REGION Network 5: Tempo total do sinal da fabrica
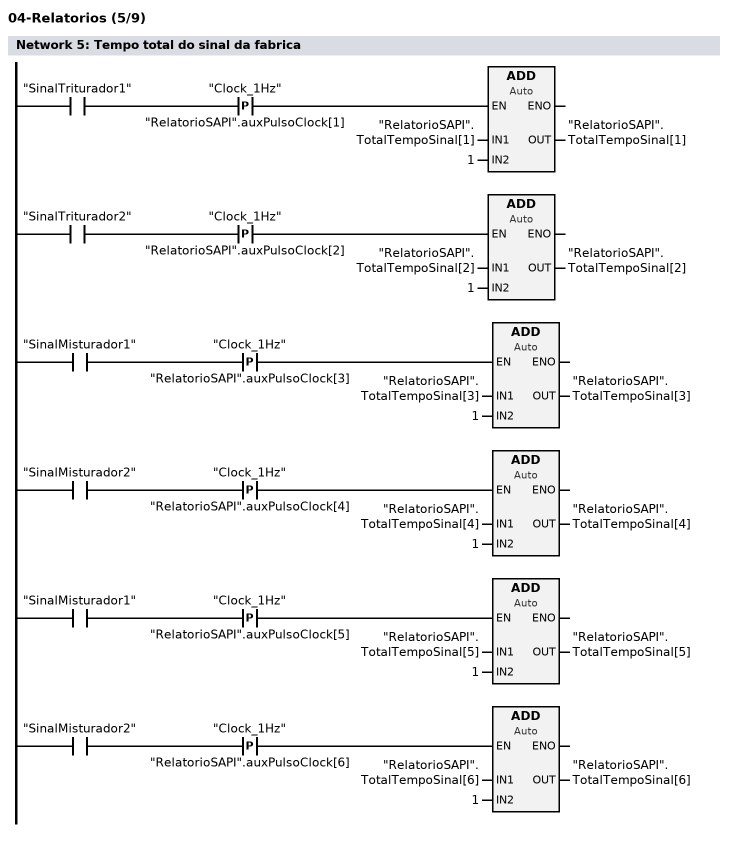
   RUNG wire#powerrail
      Contact( "SinalTriturador1" )
      P_Contact(operand := "Clock_1Hz", bit := "RelatorioSAPI".auxPulsoClock[1])
      Add(in1 := "RelatorioSAPI".TotalTempoSinal[1], in2 := 1, out => "RelatorioSAPI".TotalTempoSinal[1])
   END_RUNG
   RUNG wire#powerrail
      Contact( "SinalTriturador2" )
      P_Contact(operand := "Clock_1Hz", bit := "RelatorioSAPI".auxPulsoClock[2])
      Add(in1 := "RelatorioSAPI".TotalTempoSinal[2], in2 := 1, out => "RelatorioSAPI".TotalTempoSinal[2])
   END_RUNG
   RUNG wire#powerrail
      Contact( "SinalMisturador1" )
      P_Contact(operand := "Clock_1Hz", bit := "RelatorioSAPI".auxPulsoClock[3])
      Add(in1 := "RelatorioSAPI".TotalTempoSinal[3], in2 := 1, out => "RelatorioSAPI".TotalTempoSinal[3])
   END_RUNG
   RUNG wire#powerrail
      Contact( "SinalMisturador2" )
      P_Contact(operand := "Clock_1Hz", bit := "RelatorioSAPI".auxPulsoClock[4])
      Add(in1 := "RelatorioSAPI".TotalTempoSinal[4], in2 := 1, out => "RelatorioSAPI".TotalTempoSinal[4])
   END_RUNG
   RUNG wire#powerrail
      Contact( "SinalMisturador1" )
      P_Contact(operand := "Clock_1Hz", bit := "RelatorioSAPI".auxPulsoClock[5])
      Add(in1 := "RelatorioSAPI".TotalTempoSinal[5], in2 := 1, out => "RelatorioSAPI".TotalTempoSinal[5])
   END_RUNG
   RUNG wire#powerrail
      Contact( "SinalMisturador2" )
      P_Contact(operand := "Clock_1Hz", bit := "RelatorioSAPI".auxPulsoClock[6])
      Add(in1 := "RelatorioSAPI".TotalTempoSinal[6], in2 := 1, out => "RelatorioSAPI".TotalTempoSinal[6])
   END_RUNG
   // the same network as SCL:
   #_w1 := "SinalTriturador1" AND "Clock_1Hz" AND NOT "RelatorioSAPI".auxPulsoClock[1];   // rising edge of "Clock_1Hz"
   "RelatorioSAPI".auxPulsoClock[1] := "Clock_1Hz";
   IF #_w1 THEN "RelatorioSAPI".TotalTempoSinal[1] := "RelatorioSAPI".TotalTempoSinal[1] + 1; END_IF;
   #_w2 := "SinalTriturador2" AND "Clock_1Hz" AND NOT "RelatorioSAPI".auxPulsoClock[2];   // rising edge of "Clock_1Hz"
   "RelatorioSAPI".auxPulsoClock[2] := "Clock_1Hz";
   IF #_w2 THEN "RelatorioSAPI".TotalTempoSinal[2] := "RelatorioSAPI".TotalTempoSinal[2] + 1; END_IF;
   #_w3 := "SinalMisturador1" AND "Clock_1Hz" AND NOT "RelatorioSAPI".auxPulsoClock[3];   // rising edge of "Clock_1Hz"
   "RelatorioSAPI".auxPulsoClock[3] := "Clock_1Hz";
   IF #_w3 THEN "RelatorioSAPI".TotalTempoSinal[3] := "RelatorioSAPI".TotalTempoSinal[3] + 1; END_IF;
   #_w4 := "SinalMisturador2" AND "Clock_1Hz" AND NOT "RelatorioSAPI".auxPulsoClock[4];   // rising edge of "Clock_1Hz"
   "RelatorioSAPI".auxPulsoClock[4] := "Clock_1Hz";
   IF #_w4 THEN "RelatorioSAPI".TotalTempoSinal[4] := "RelatorioSAPI".TotalTempoSinal[4] + 1; END_IF;
   #_w5 := "SinalMisturador1" AND "Clock_1Hz" AND NOT "RelatorioSAPI".auxPulsoClock[5];   // rising edge of "Clock_1Hz"
   "RelatorioSAPI".auxPulsoClock[5] := "Clock_1Hz";
   IF #_w5 THEN "RelatorioSAPI".TotalTempoSinal[5] := "RelatorioSAPI".TotalTempoSinal[5] + 1; END_IF;
   #_w6 := "SinalMisturador2" AND "Clock_1Hz" AND NOT "RelatorioSAPI".auxPulsoClock[6];   // rising edge of "Clock_1Hz"
   "RelatorioSAPI".auxPulsoClock[6] := "Clock_1Hz";
   IF #_w6 THEN "RelatorioSAPI".TotalTempoSinal[6] := "RelatorioSAPI".TotalTempoSinal[6] + 1; END_IF;
END_REGION

REGION Network 6: Quantidade acionamentos sinal fabrica
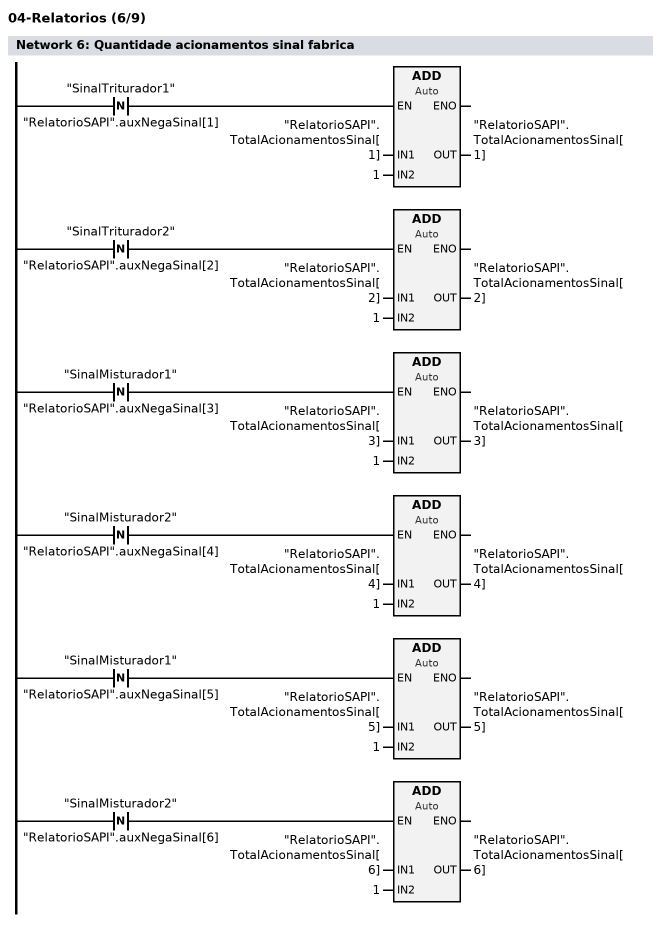
   RUNG wire#powerrail
      N_Contact(operand := "SinalTriturador1", bit := "RelatorioSAPI".auxNegaSinal[1])
      Add(in1 := "RelatorioSAPI".TotalAcionamentosSinal[1], in2 := 1, out => "RelatorioSAPI".TotalAcionamentosSinal[1])
   END_RUNG
   RUNG wire#powerrail
      N_Contact(operand := "SinalTriturador2", bit := "RelatorioSAPI".auxNegaSinal[2])
      Add(in1 := "RelatorioSAPI".TotalAcionamentosSinal[2], in2 := 1, out => "RelatorioSAPI".TotalAcionamentosSinal[2])
   END_RUNG
   RUNG wire#powerrail
      N_Contact(operand := "SinalMisturador1", bit := "RelatorioSAPI".auxNegaSinal[3])
      Add(in1 := "RelatorioSAPI".TotalAcionamentosSinal[3], in2 := 1, out => "RelatorioSAPI".TotalAcionamentosSinal[3])
   END_RUNG
   RUNG wire#powerrail
      N_Contact(operand := "SinalMisturador2", bit := "RelatorioSAPI".auxNegaSinal[4])
      Add(in1 := "RelatorioSAPI".TotalAcionamentosSinal[4], in2 := 1, out => "RelatorioSAPI".TotalAcionamentosSinal[4])
   END_RUNG
   RUNG wire#powerrail
      N_Contact(operand := "SinalMisturador1", bit := "RelatorioSAPI".auxNegaSinal[5])
      Add(in1 := "RelatorioSAPI".TotalAcionamentosSinal[5], in2 := 1, out => "RelatorioSAPI".TotalAcionamentosSinal[5])
   END_RUNG
   RUNG wire#powerrail
      N_Contact(operand := "SinalMisturador2", bit := "RelatorioSAPI".auxNegaSinal[6])
      Add(in1 := "RelatorioSAPI".TotalAcionamentosSinal[6], in2 := 1, out => "RelatorioSAPI".TotalAcionamentosSinal[6])
   END_RUNG
   // the same network as SCL:
   #_w1 := NOT "SinalTriturador1" AND "RelatorioSAPI".auxNegaSinal[1];   // falling edge of "SinalTriturador1"
   "RelatorioSAPI".auxNegaSinal[1] := "SinalTriturador1";
   IF #_w1 THEN
       "RelatorioSAPI".TotalAcionamentosSinal[1] := "RelatorioSAPI".TotalAcionamentosSinal[1] + 1;
   END_IF;
   #_w2 := NOT "SinalTriturador2" AND "RelatorioSAPI".auxNegaSinal[2];   // falling edge of "SinalTriturador2"
   "RelatorioSAPI".auxNegaSinal[2] := "SinalTriturador2";
   IF #_w2 THEN
       "RelatorioSAPI".TotalAcionamentosSinal[2] := "RelatorioSAPI".TotalAcionamentosSinal[2] + 1;
   END_IF;
   #_w3 := NOT "SinalMisturador1" AND "RelatorioSAPI".auxNegaSinal[3];   // falling edge of "SinalMisturador1"
   "RelatorioSAPI".auxNegaSinal[3] := "SinalMisturador1";
   IF #_w3 THEN
       "RelatorioSAPI".TotalAcionamentosSinal[3] := "RelatorioSAPI".TotalAcionamentosSinal[3] + 1;
   END_IF;
   #_w4 := NOT "SinalMisturador2" AND "RelatorioSAPI".auxNegaSinal[4];   // falling edge of "SinalMisturador2"
   "RelatorioSAPI".auxNegaSinal[4] := "SinalMisturador2";
   IF #_w4 THEN
       "RelatorioSAPI".TotalAcionamentosSinal[4] := "RelatorioSAPI".TotalAcionamentosSinal[4] + 1;
   END_IF;
   #_w5 := NOT "SinalMisturador1" AND "RelatorioSAPI".auxNegaSinal[5];   // falling edge of "SinalMisturador1"
   "RelatorioSAPI".auxNegaSinal[5] := "SinalMisturador1";
   IF #_w5 THEN
       "RelatorioSAPI".TotalAcionamentosSinal[5] := "RelatorioSAPI".TotalAcionamentosSinal[5] + 1;
   END_IF;
   #_w6 := NOT "SinalMisturador2" AND "RelatorioSAPI".auxNegaSinal[6];   // falling edge of "SinalMisturador2"
   "RelatorioSAPI".auxNegaSinal[6] := "SinalMisturador2";
   IF #_w6 THEN
       "RelatorioSAPI".TotalAcionamentosSinal[6] := "RelatorioSAPI".TotalAcionamentosSinal[6] + 1;
   END_IF;
END_REGION

REGION Network 7: Quantidade acionamentos bombas
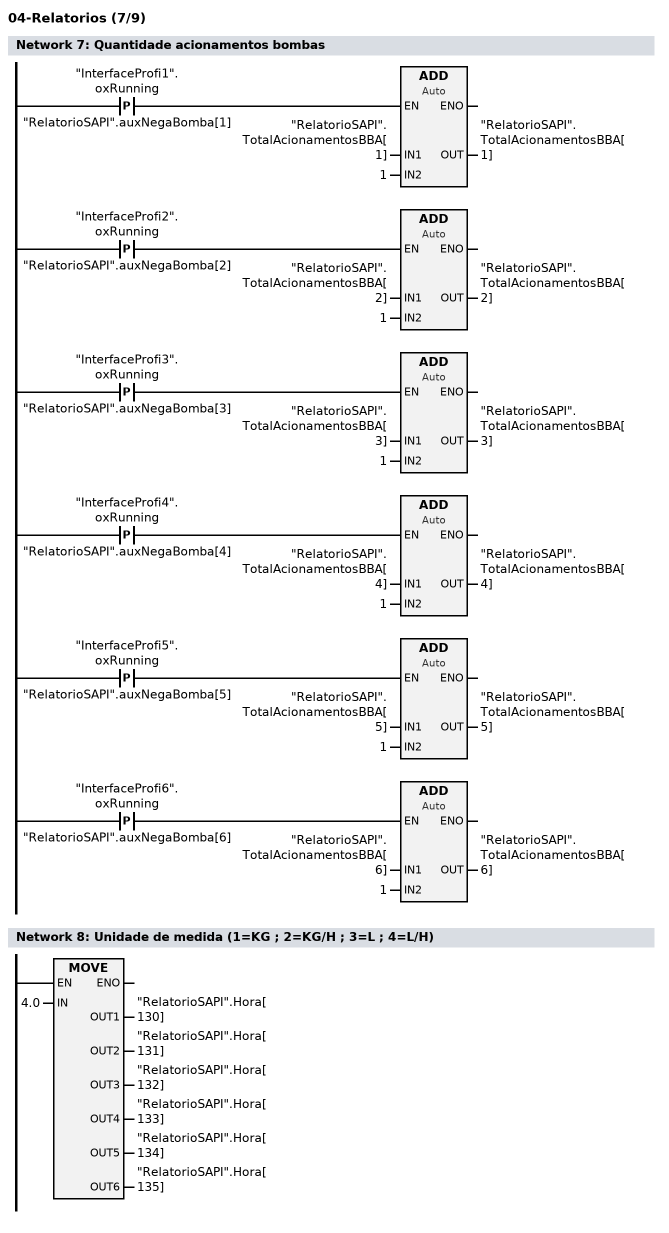
   RUNG wire#powerrail
      P_Contact(operand := "InterfaceProfi1".oxRunning, bit := "RelatorioSAPI".auxNegaBomba[1])
      Add(in1 := "RelatorioSAPI".TotalAcionamentosBBA[1], in2 := 1, out => "RelatorioSAPI".TotalAcionamentosBBA[1])
   END_RUNG
   RUNG wire#powerrail
      P_Contact(operand := "InterfaceProfi2".oxRunning, bit := "RelatorioSAPI".auxNegaBomba[2])
      Add(in1 := "RelatorioSAPI".TotalAcionamentosBBA[2], in2 := 1, out => "RelatorioSAPI".TotalAcionamentosBBA[2])
   END_RUNG
   RUNG wire#powerrail
      P_Contact(operand := "InterfaceProfi3".oxRunning, bit := "RelatorioSAPI".auxNegaBomba[3])
      Add(in1 := "RelatorioSAPI".TotalAcionamentosBBA[3], in2 := 1, out => "RelatorioSAPI".TotalAcionamentosBBA[3])
   END_RUNG
   RUNG wire#powerrail
      P_Contact(operand := "InterfaceProfi4".oxRunning, bit := "RelatorioSAPI".auxNegaBomba[4])
      Add(in1 := "RelatorioSAPI".TotalAcionamentosBBA[4], in2 := 1, out => "RelatorioSAPI".TotalAcionamentosBBA[4])
   END_RUNG
   RUNG wire#powerrail
      P_Contact(operand := "InterfaceProfi5".oxRunning, bit := "RelatorioSAPI".auxNegaBomba[5])
      Add(in1 := "RelatorioSAPI".TotalAcionamentosBBA[5], in2 := 1, out => "RelatorioSAPI".TotalAcionamentosBBA[5])
   END_RUNG
   RUNG wire#powerrail
      P_Contact(operand := "InterfaceProfi6".oxRunning, bit := "RelatorioSAPI".auxNegaBomba[6])
      Add(in1 := "RelatorioSAPI".TotalAcionamentosBBA[6], in2 := 1, out => "RelatorioSAPI".TotalAcionamentosBBA[6])
   END_RUNG
   // the same network as SCL:
   #_w1 := "InterfaceProfi1".oxRunning AND NOT "RelatorioSAPI".auxNegaBomba[1];   // rising edge of "InterfaceProfi1".oxRunning
   "RelatorioSAPI".auxNegaBomba[1] := "InterfaceProfi1".oxRunning;
   IF #_w1 THEN
       "RelatorioSAPI".TotalAcionamentosBBA[1] := "RelatorioSAPI".TotalAcionamentosBBA[1] + 1;
   END_IF;
   #_w2 := "InterfaceProfi2".oxRunning AND NOT "RelatorioSAPI".auxNegaBomba[2];   // rising edge of "InterfaceProfi2".oxRunning
   "RelatorioSAPI".auxNegaBomba[2] := "InterfaceProfi2".oxRunning;
   IF #_w2 THEN
       "RelatorioSAPI".TotalAcionamentosBBA[2] := "RelatorioSAPI".TotalAcionamentosBBA[2] + 1;
   END_IF;
   #_w3 := "InterfaceProfi3".oxRunning AND NOT "RelatorioSAPI".auxNegaBomba[3];   // rising edge of "InterfaceProfi3".oxRunning
   "RelatorioSAPI".auxNegaBomba[3] := "InterfaceProfi3".oxRunning;
   IF #_w3 THEN
       "RelatorioSAPI".TotalAcionamentosBBA[3] := "RelatorioSAPI".TotalAcionamentosBBA[3] + 1;
   END_IF;
   #_w4 := "InterfaceProfi4".oxRunning AND NOT "RelatorioSAPI".auxNegaBomba[4];   // rising edge of "InterfaceProfi4".oxRunning
   "RelatorioSAPI".auxNegaBomba[4] := "InterfaceProfi4".oxRunning;
   IF #_w4 THEN
       "RelatorioSAPI".TotalAcionamentosBBA[4] := "RelatorioSAPI".TotalAcionamentosBBA[4] + 1;
   END_IF;
   #_w5 := "InterfaceProfi5".oxRunning AND NOT "RelatorioSAPI".auxNegaBomba[5];   // rising edge of "InterfaceProfi5".oxRunning
   "RelatorioSAPI".auxNegaBomba[5] := "InterfaceProfi5".oxRunning;
   IF #_w5 THEN
       "RelatorioSAPI".TotalAcionamentosBBA[5] := "RelatorioSAPI".TotalAcionamentosBBA[5] + 1;
   END_IF;
   #_w6 := "InterfaceProfi6".oxRunning AND NOT "RelatorioSAPI".auxNegaBomba[6];   // rising edge of "InterfaceProfi6".oxRunning
   "RelatorioSAPI".auxNegaBomba[6] := "InterfaceProfi6".oxRunning;
   IF #_w6 THEN
       "RelatorioSAPI".TotalAcionamentosBBA[6] := "RelatorioSAPI".TotalAcionamentosBBA[6] + 1;
   END_IF;
END_REGION

REGION Network 8: Unidade de medida (1=KG ; 2=KG/H ; 3=L ; 4=L/H)
   RUNG wire#powerrail
      Move(in := 4.0, out1 => "RelatorioSAPI".Hora[130], out2 => "RelatorioSAPI".Hora[131], out3 => "RelatorioSAPI".Hora[132], out4 => "RelatorioSAPI".Hora[133], out5 => "RelatorioSAPI".Hora[134], out6 => "RelatorioSAPI".Hora[135])
   END_RUNG
   // the same network as SCL:
   "RelatorioSAPI".Hora[130] := 4.0;
   "RelatorioSAPI".Hora[131] := 4.0;
   "RelatorioSAPI".Hora[132] := 4.0;
   "RelatorioSAPI".Hora[133] := 4.0;
   "RelatorioSAPI".Hora[134] := 4.0;
   "RelatorioSAPI".Hora[135] := 4.0;
END_REGION

REGION Network 9: NOME DA BOMBA
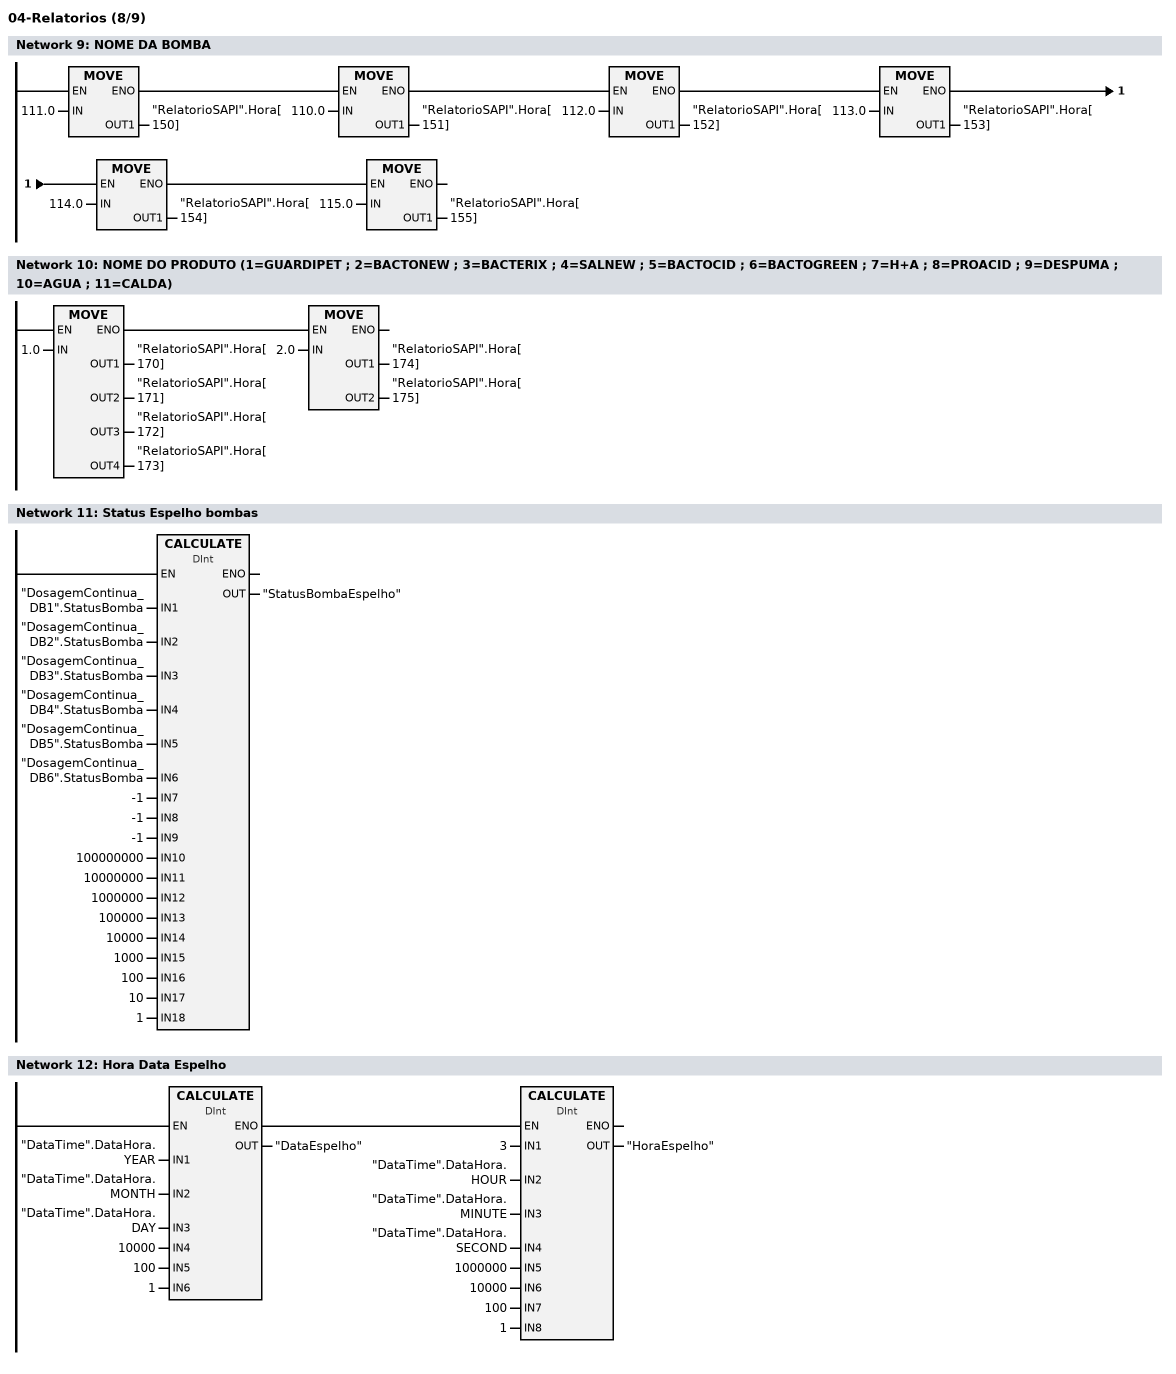
   RUNG wire#powerrail
      Move(in := 111.0, out1 => "RelatorioSAPI".Hora[150])
      Move(in := 110.0, out1 => "RelatorioSAPI".Hora[151])
      Move(in := 112.0, out1 => "RelatorioSAPI".Hora[152])
      Move(in := 113.0, out1 => "RelatorioSAPI".Hora[153])
      Move(in := 114.0, out1 => "RelatorioSAPI".Hora[154])
      Move(in := 115.0, out1 => "RelatorioSAPI".Hora[155])
   END_RUNG
   // the same network as SCL:
   "RelatorioSAPI".Hora[150] := 111.0;
   "RelatorioSAPI".Hora[151] := 110.0;
   "RelatorioSAPI".Hora[152] := 112.0;
   "RelatorioSAPI".Hora[153] := 113.0;
   "RelatorioSAPI".Hora[154] := 114.0;
   "RelatorioSAPI".Hora[155] := 115.0;
END_REGION

REGION Network 10: NOME DO PRODUTO (1=GUARDIPET ; 2=BACTONEW ; 3=BACTERIX ; 4=SALNEW ; 5=BACTOCID ; 6=BACTOGREEN ; 7=H+A ; 8=PROACID ; 9=DESPUMA ; 10=AGUA ; 11=CALDA)
   RUNG wire#powerrail
      Move(in := 1.0, out1 => "RelatorioSAPI".Hora[170], out2 => "RelatorioSAPI".Hora[171], out3 => "RelatorioSAPI".Hora[172], out4 => "RelatorioSAPI".Hora[173])
      Move(in := 2.0, out1 => "RelatorioSAPI".Hora[174], out2 => "RelatorioSAPI".Hora[175])
   END_RUNG
   // the same network as SCL:
   "RelatorioSAPI".Hora[170] := 1.0;
   "RelatorioSAPI".Hora[171] := 1.0;
   "RelatorioSAPI".Hora[172] := 1.0;
   "RelatorioSAPI".Hora[173] := 1.0;
   "RelatorioSAPI".Hora[174] := 2.0;
   "RelatorioSAPI".Hora[175] := 2.0;
END_REGION

REGION Network 11: Status Espelho bombas
   RUNG wire#powerrail
      { S7_Templates := "SrcType := DInt"; S7_Expression := "(((IN18+IN1) * IN10) + ((IN18+IN2) * IN11) + ((IN18+IN3) * IN12) + ((IN18+IN4) * IN13) + ((IN18+IN5) * IN14) + ((IN18+IN6) * IN15) + ((IN18+IN7) * IN16) + ((IN18+IN8) * IN17) + ((IN18+IN9) * IN18))" } Calculate(in1 := "DosagemContinua_DB1".StatusBomba, in2 := "DosagemContinua_DB2".StatusBomba, in3 := "DosagemContinua_DB3".StatusBomba, in4 := "DosagemContinua_DB4".StatusBomba, in5 := "DosagemContinua_DB5".StatusBomba, in6 := "DosagemContinua_DB6".StatusBomba, in7 := -1, in8 := -1, in9 := -1, in10 := 100000000, in11 := 10000000, in12 := 1000000, in13 := 100000, in14 := 10000, in15 := 1000, in16 := 100, in17 := 10, in18 := 1, out => "StatusBombaEspelho")
   END_RUNG
   // the same network as SCL:
   "StatusBombaEspelho" := (((1+"DosagemContinua_DB1".StatusBomba) * 100000000) + ((1+"DosagemContinua_DB2".StatusBomba) * 10000000) + ((1+"DosagemContinua_DB3".StatusBomba) * 1000000) + ((1+"DosagemContinua_DB4".StatusBomba) * 100000) + ((1+"DosagemContinua_DB5".StatusBomba) * 10000) + ((1+"DosagemContinua_DB6".StatusBomba) * 1000) + ((1+(-1)) * 100) + ((1+(-1)) * 10) + ((1+(-1)) * 1));
END_REGION

REGION Network 12: Hora Data Espelho
   RUNG wire#powerrail
      { S7_Templates := "SrcType := DInt"; S7_Expression := "((IN1 * IN4) + (IN2 * IN5) + (IN3 * IN6))" } Calculate(in1 := "DataTime".DataHora.YEAR, in2 := "DataTime".DataHora.MONTH, in3 := "DataTime".DataHora.DAY, in4 := 10000, in5 := 100, in6 := 1, out => "DataEspelho")
      { S7_Templates := "SrcType := DInt"; S7_Expression := "((IN1 * IN5) + (IN2 * IN6) + (IN3 * IN7) + (IN4 * IN8))" } Calculate(in1 := 3, in2 := "DataTime".DataHora.HOUR, in3 := "DataTime".DataHora.MINUTE, in4 := "DataTime".DataHora.SECOND, in5 := 1000000, in6 := 10000, in7 := 100, in8 := 1, out => "HoraEspelho")
   END_RUNG
   // the same network as SCL:
   "DataEspelho" := (("DataTime".DataHora.YEAR * 10000) + ("DataTime".DataHora.MONTH * 100) + ("DataTime".DataHora.DAY * 1));
   "HoraEspelho" := ((3 * 1000000) + ("DataTime".DataHora.HOUR * 10000) + ("DataTime".DataHora.MINUTE * 100) + ("DataTime".DataHora.SECOND * 1));
END_REGION

REGION Network 13: RELATORIO SAPI
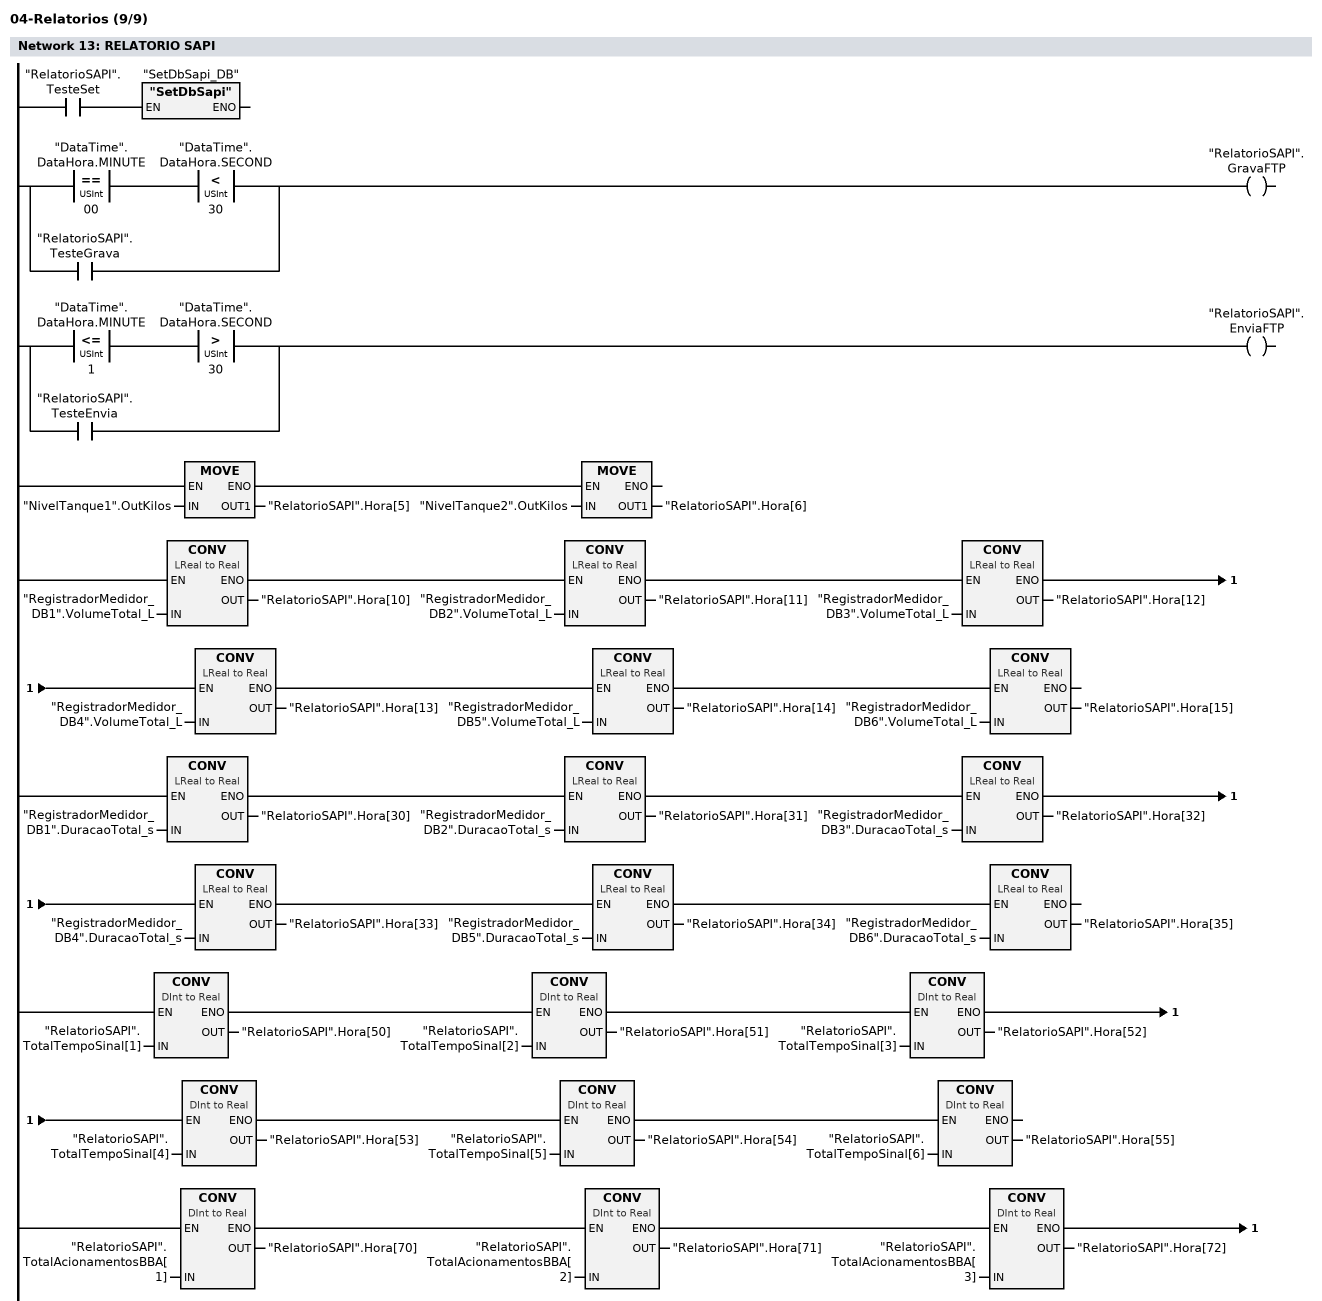
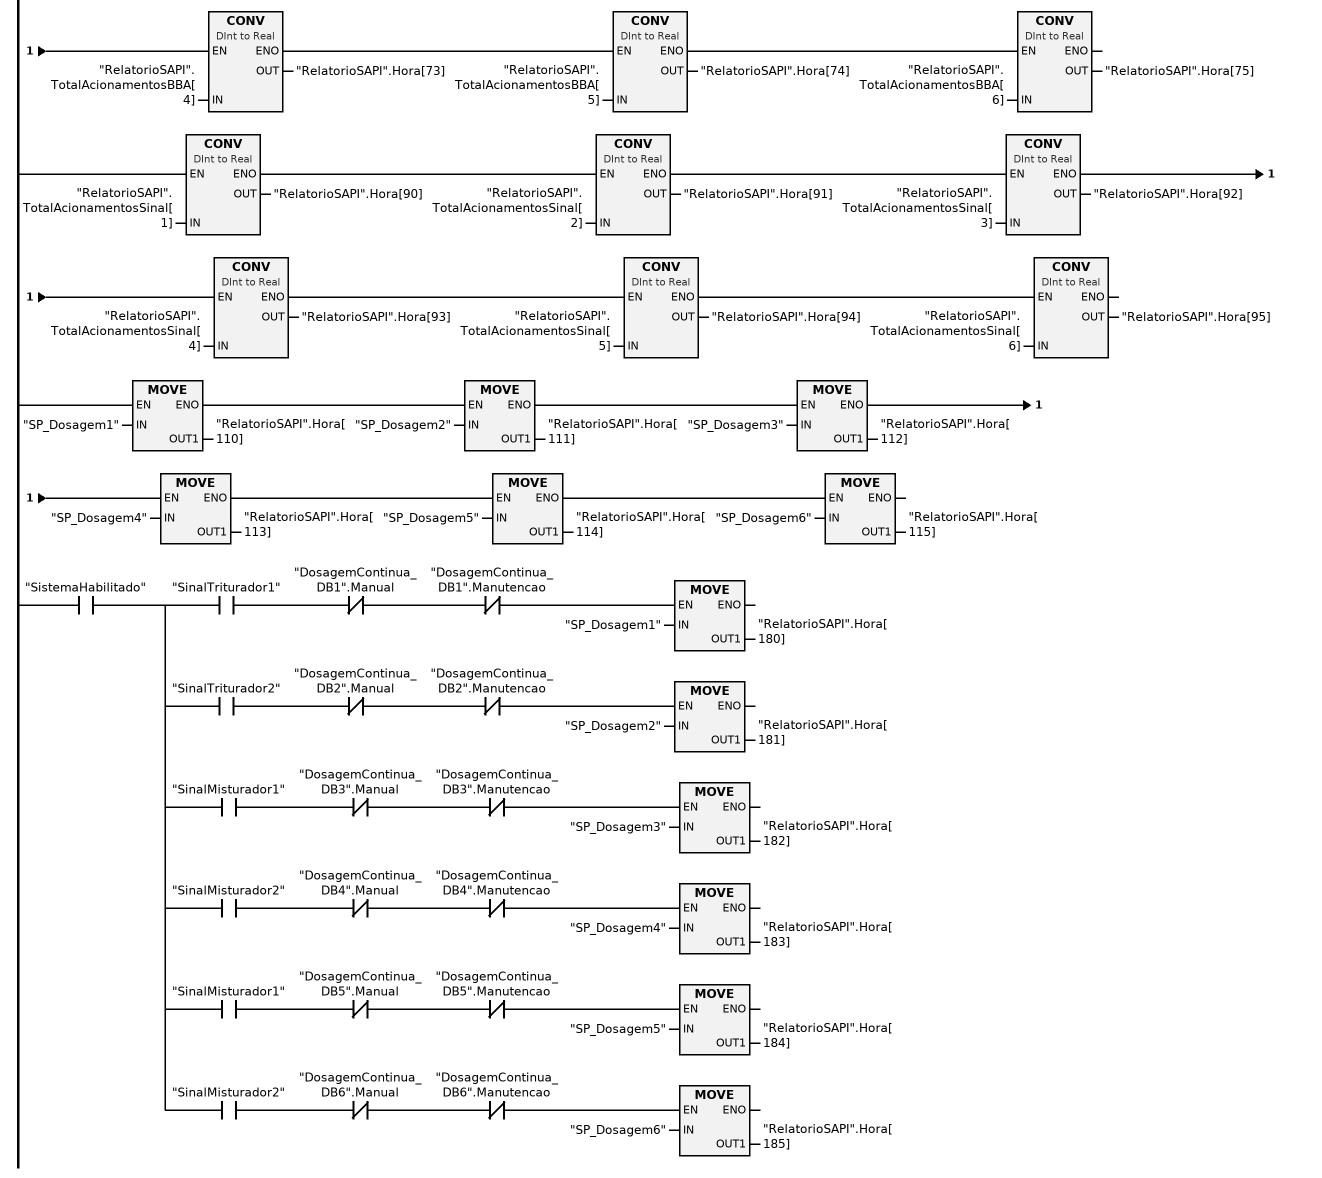
   RUNG wire#powerrail
      Contact( "RelatorioSAPI".TesteSet )
      "SetDbSapi_DB"()
   END_RUNG
   RUNG wire#powerrail
      { S7_Templates := "SrcType := USInt" } EQ_Contact(in1 := "DataTime".DataHora.MINUTE, in2 := 00)
      { S7_Templates := "SrcType := USInt" } LT_Contact(in1 := "DataTime".DataHora.SECOND, in2 := 30)
      wire#w1
      Coil( "RelatorioSAPI".GravaFTP )
   END_RUNG
   RUNG wire#powerrail
      Contact( "RelatorioSAPI".TesteGrava )
   END_RUNG wire#w1
   RUNG wire#powerrail
      { S7_Templates := "SrcType := USInt" } LE_Contact(in1 := "DataTime".DataHora.MINUTE, in2 := 1)
      { S7_Templates := "SrcType := USInt" } GT_Contact(in1 := "DataTime".DataHora.SECOND, in2 := 30)
      wire#w2
      Coil( "RelatorioSAPI".EnviaFTP )
   END_RUNG
   RUNG wire#powerrail
      Contact( "RelatorioSAPI".TesteEnvia )
   END_RUNG wire#w2
   RUNG wire#powerrail
      Move(in := "NivelTanque1".OutKilos, out1 => "RelatorioSAPI".Hora[5])
      Move(in := "NivelTanque2".OutKilos, out1 => "RelatorioSAPI".Hora[6])
   END_RUNG
   RUNG wire#powerrail
      { S7_Templates := "[SrcType := LReal, DestType := Real]" } Convert(in := "RegistradorMedidor_DB1".VolumeTotal_L, out => "RelatorioSAPI".Hora[10])
      { S7_Templates := "[SrcType := LReal, DestType := Real]" } Convert(in := "RegistradorMedidor_DB2".VolumeTotal_L, out => "RelatorioSAPI".Hora[11])
      { S7_Templates := "[SrcType := LReal, DestType := Real]" } Convert(in := "RegistradorMedidor_DB3".VolumeTotal_L, out => "RelatorioSAPI".Hora[12])
      { S7_Templates := "[SrcType := LReal, DestType := Real]" } Convert(in := "RegistradorMedidor_DB4".VolumeTotal_L, out => "RelatorioSAPI".Hora[13])
      { S7_Templates := "[SrcType := LReal, DestType := Real]" } Convert(in := "RegistradorMedidor_DB5".VolumeTotal_L, out => "RelatorioSAPI".Hora[14])
      { S7_Templates := "[SrcType := LReal, DestType := Real]" } Convert(in := "RegistradorMedidor_DB6".VolumeTotal_L, out => "RelatorioSAPI".Hora[15])
   END_RUNG
   RUNG wire#powerrail
      { S7_Templates := "[SrcType := LReal, DestType := Real]" } Convert(in := "RegistradorMedidor_DB1".DuracaoTotal_s, out => "RelatorioSAPI".Hora[30])
      { S7_Templates := "[SrcType := LReal, DestType := Real]" } Convert(in := "RegistradorMedidor_DB2".DuracaoTotal_s, out => "RelatorioSAPI".Hora[31])
      { S7_Templates := "[SrcType := LReal, DestType := Real]" } Convert(in := "RegistradorMedidor_DB3".DuracaoTotal_s, out => "RelatorioSAPI".Hora[32])
      { S7_Templates := "[SrcType := LReal, DestType := Real]" } Convert(in := "RegistradorMedidor_DB4".DuracaoTotal_s, out => "RelatorioSAPI".Hora[33])
      { S7_Templates := "[SrcType := LReal, DestType := Real]" } Convert(in := "RegistradorMedidor_DB5".DuracaoTotal_s, out => "RelatorioSAPI".Hora[34])
      { S7_Templates := "[SrcType := LReal, DestType := Real]" } Convert(in := "RegistradorMedidor_DB6".DuracaoTotal_s, out => "RelatorioSAPI".Hora[35])
   END_RUNG
   RUNG wire#powerrail
      { S7_Templates := "[SrcType := DInt, DestType := Real]" } Convert(in := "RelatorioSAPI".TotalTempoSinal[1], out => "RelatorioSAPI".Hora[50])
      { S7_Templates := "[SrcType := DInt, DestType := Real]" } Convert(in := "RelatorioSAPI".TotalTempoSinal[2], out => "RelatorioSAPI".Hora[51])
      { S7_Templates := "[SrcType := DInt, DestType := Real]" } Convert(in := "RelatorioSAPI".TotalTempoSinal[3], out => "RelatorioSAPI".Hora[52])
      { S7_Templates := "[SrcType := DInt, DestType := Real]" } Convert(in := "RelatorioSAPI".TotalTempoSinal[4], out => "RelatorioSAPI".Hora[53])
      { S7_Templates := "[SrcType := DInt, DestType := Real]" } Convert(in := "RelatorioSAPI".TotalTempoSinal[5], out => "RelatorioSAPI".Hora[54])
      { S7_Templates := "[SrcType := DInt, DestType := Real]" } Convert(in := "RelatorioSAPI".TotalTempoSinal[6], out => "RelatorioSAPI".Hora[55])
   END_RUNG
   RUNG wire#powerrail
      { S7_Templates := "[SrcType := DInt, DestType := Real]" } Convert(in := "RelatorioSAPI".TotalAcionamentosBBA[1], out => "RelatorioSAPI".Hora[70])
      { S7_Templates := "[SrcType := DInt, DestType := Real]" } Convert(in := "RelatorioSAPI".TotalAcionamentosBBA[2], out => "RelatorioSAPI".Hora[71])
      { S7_Templates := "[SrcType := DInt, DestType := Real]" } Convert(in := "RelatorioSAPI".TotalAcionamentosBBA[3], out => "RelatorioSAPI".Hora[72])
      { S7_Templates := "[SrcType := DInt, DestType := Real]" } Convert(in := "RelatorioSAPI".TotalAcionamentosBBA[4], out => "RelatorioSAPI".Hora[73])
      { S7_Templates := "[SrcType := DInt, DestType := Real]" } Convert(in := "RelatorioSAPI".TotalAcionamentosBBA[5], out => "RelatorioSAPI".Hora[74])
      { S7_Templates := "[SrcType := DInt, DestType := Real]" } Convert(in := "RelatorioSAPI".TotalAcionamentosBBA[6], out => "RelatorioSAPI".Hora[75])
   END_RUNG
   RUNG wire#powerrail
      { S7_Templates := "[SrcType := DInt, DestType := Real]" } Convert(in := "RelatorioSAPI".TotalAcionamentosSinal[1], out => "RelatorioSAPI".Hora[90])
      { S7_Templates := "[SrcType := DInt, DestType := Real]" } Convert(in := "RelatorioSAPI".TotalAcionamentosSinal[2], out => "RelatorioSAPI".Hora[91])
      { S7_Templates := "[SrcType := DInt, DestType := Real]" } Convert(in := "RelatorioSAPI".TotalAcionamentosSinal[3], out => "RelatorioSAPI".Hora[92])
      { S7_Templates := "[SrcType := DInt, DestType := Real]" } Convert(in := "RelatorioSAPI".TotalAcionamentosSinal[4], out => "RelatorioSAPI".Hora[93])
      { S7_Templates := "[SrcType := DInt, DestType := Real]" } Convert(in := "RelatorioSAPI".TotalAcionamentosSinal[5], out => "RelatorioSAPI".Hora[94])
      { S7_Templates := "[SrcType := DInt, DestType := Real]" } Convert(in := "RelatorioSAPI".TotalAcionamentosSinal[6], out => "RelatorioSAPI".Hora[95])
   END_RUNG
   RUNG wire#powerrail
      Move(in := "SP_Dosagem1", out1 => "RelatorioSAPI".Hora[110])
      Move(in := "SP_Dosagem2", out1 => "RelatorioSAPI".Hora[111])
      Move(in := "SP_Dosagem3", out1 => "RelatorioSAPI".Hora[112])
      Move(in := "SP_Dosagem4", out1 => "RelatorioSAPI".Hora[113])
      Move(in := "SP_Dosagem5", out1 => "RelatorioSAPI".Hora[114])
      Move(in := "SP_Dosagem6", out1 => "RelatorioSAPI".Hora[115])
   END_RUNG
   RUNG wire#powerrail
      Contact( "SistemaHabilitado" )
      wire#w3
      Contact( "SinalTriturador1" )
      I_Contact( "DosagemContinua_DB1".Manual )
      I_Contact( "DosagemContinua_DB1".Manutencao )
      Move(in := "SP_Dosagem1", out1 => "RelatorioSAPI".Hora[180])
   END_RUNG
   RUNG wire#w3
      Contact( "SinalTriturador2" )
      I_Contact( "DosagemContinua_DB2".Manual )
      I_Contact( "DosagemContinua_DB2".Manutencao )
      Move(in := "SP_Dosagem2", out1 => "RelatorioSAPI".Hora[181])
   END_RUNG
   RUNG wire#w3
      Contact( "SinalMisturador1" )
      I_Contact( "DosagemContinua_DB3".Manual )
      I_Contact( "DosagemContinua_DB3".Manutencao )
      Move(in := "SP_Dosagem3", out1 => "RelatorioSAPI".Hora[182])
   END_RUNG
   RUNG wire#w3
      Contact( "SinalMisturador2" )
      I_Contact( "DosagemContinua_DB4".Manual )
      I_Contact( "DosagemContinua_DB4".Manutencao )
      Move(in := "SP_Dosagem4", out1 => "RelatorioSAPI".Hora[183])
   END_RUNG
   RUNG wire#w3
      Contact( "SinalMisturador1" )
      I_Contact( "DosagemContinua_DB5".Manual )
      I_Contact( "DosagemContinua_DB5".Manutencao )
      Move(in := "SP_Dosagem5", out1 => "RelatorioSAPI".Hora[184])
   END_RUNG
   RUNG wire#w3
      Contact( "SinalMisturador2" )
      I_Contact( "DosagemContinua_DB6".Manual )
      I_Contact( "DosagemContinua_DB6".Manutencao )
      Move(in := "SP_Dosagem6", out1 => "RelatorioSAPI".Hora[185])
   END_RUNG
   // the same network as SCL:
   IF "RelatorioSAPI".TesteSet THEN
       "SetDbSapi_DB"();   // "SetDbSapi"
   END_IF;
   "RelatorioSAPI".GravaFTP := (("DataTime".DataHora.MINUTE = 00) AND ("DataTime".DataHora.SECOND < 30)) OR "RelatorioSAPI".TesteGrava;
   "RelatorioSAPI".EnviaFTP := (("DataTime".DataHora.MINUTE <= 1) AND ("DataTime".DataHora.SECOND > 30)) OR "RelatorioSAPI".TesteEnvia;
   "RelatorioSAPI".Hora[5] := "NivelTanque1".OutKilos;
   "RelatorioSAPI".Hora[6] := "NivelTanque2".OutKilos;
   "RelatorioSAPI".Hora[10] := LREAL_TO_REAL("RegistradorMedidor_DB1".VolumeTotal_L);
   "RelatorioSAPI".Hora[11] := LREAL_TO_REAL("RegistradorMedidor_DB2".VolumeTotal_L);
   "RelatorioSAPI".Hora[12] := LREAL_TO_REAL("RegistradorMedidor_DB3".VolumeTotal_L);
   "RelatorioSAPI".Hora[13] := LREAL_TO_REAL("RegistradorMedidor_DB4".VolumeTotal_L);
   "RelatorioSAPI".Hora[14] := LREAL_TO_REAL("RegistradorMedidor_DB5".VolumeTotal_L);
   "RelatorioSAPI".Hora[15] := LREAL_TO_REAL("RegistradorMedidor_DB6".VolumeTotal_L);
   "RelatorioSAPI".Hora[30] := LREAL_TO_REAL("RegistradorMedidor_DB1".DuracaoTotal_s);
   "RelatorioSAPI".Hora[31] := LREAL_TO_REAL("RegistradorMedidor_DB2".DuracaoTotal_s);
   "RelatorioSAPI".Hora[32] := LREAL_TO_REAL("RegistradorMedidor_DB3".DuracaoTotal_s);
   "RelatorioSAPI".Hora[33] := LREAL_TO_REAL("RegistradorMedidor_DB4".DuracaoTotal_s);
   "RelatorioSAPI".Hora[34] := LREAL_TO_REAL("RegistradorMedidor_DB5".DuracaoTotal_s);
   "RelatorioSAPI".Hora[35] := LREAL_TO_REAL("RegistradorMedidor_DB6".DuracaoTotal_s);
   "RelatorioSAPI".Hora[50] := DINT_TO_REAL("RelatorioSAPI".TotalTempoSinal[1]);
   "RelatorioSAPI".Hora[51] := DINT_TO_REAL("RelatorioSAPI".TotalTempoSinal[2]);
   "RelatorioSAPI".Hora[52] := DINT_TO_REAL("RelatorioSAPI".TotalTempoSinal[3]);
   "RelatorioSAPI".Hora[53] := DINT_TO_REAL("RelatorioSAPI".TotalTempoSinal[4]);
   "RelatorioSAPI".Hora[54] := DINT_TO_REAL("RelatorioSAPI".TotalTempoSinal[5]);
   "RelatorioSAPI".Hora[55] := DINT_TO_REAL("RelatorioSAPI".TotalTempoSinal[6]);
   "RelatorioSAPI".Hora[70] := DINT_TO_REAL("RelatorioSAPI".TotalAcionamentosBBA[1]);
   "RelatorioSAPI".Hora[71] := DINT_TO_REAL("RelatorioSAPI".TotalAcionamentosBBA[2]);
   "RelatorioSAPI".Hora[72] := DINT_TO_REAL("RelatorioSAPI".TotalAcionamentosBBA[3]);
   "RelatorioSAPI".Hora[73] := DINT_TO_REAL("RelatorioSAPI".TotalAcionamentosBBA[4]);
   "RelatorioSAPI".Hora[74] := DINT_TO_REAL("RelatorioSAPI".TotalAcionamentosBBA[5]);
   "RelatorioSAPI".Hora[75] := DINT_TO_REAL("RelatorioSAPI".TotalAcionamentosBBA[6]);
   "RelatorioSAPI".Hora[90] := DINT_TO_REAL("RelatorioSAPI".TotalAcionamentosSinal[1]);
   "RelatorioSAPI".Hora[91] := DINT_TO_REAL("RelatorioSAPI".TotalAcionamentosSinal[2]);
   "RelatorioSAPI".Hora[92] := DINT_TO_REAL("RelatorioSAPI".TotalAcionamentosSinal[3]);
   "RelatorioSAPI".Hora[93] := DINT_TO_REAL("RelatorioSAPI".TotalAcionamentosSinal[4]);
   "RelatorioSAPI".Hora[94] := DINT_TO_REAL("RelatorioSAPI".TotalAcionamentosSinal[5]);
   "RelatorioSAPI".Hora[95] := DINT_TO_REAL("RelatorioSAPI".TotalAcionamentosSinal[6]);
   "RelatorioSAPI".Hora[110] := "SP_Dosagem1";
   "RelatorioSAPI".Hora[111] := "SP_Dosagem2";
   "RelatorioSAPI".Hora[112] := "SP_Dosagem3";
   "RelatorioSAPI".Hora[113] := "SP_Dosagem4";
   "RelatorioSAPI".Hora[114] := "SP_Dosagem5";
   "RelatorioSAPI".Hora[115] := "SP_Dosagem6";
   IF "SistemaHabilitado" AND "SinalTriturador1" AND NOT "DosagemContinua_DB1".Manual AND NOT "DosagemContinua_DB1".Manutencao THEN
       "RelatorioSAPI".Hora[180] := "SP_Dosagem1";
   END_IF;
   IF "SistemaHabilitado" AND "SinalTriturador2" AND NOT "DosagemContinua_DB2".Manual AND NOT "DosagemContinua_DB2".Manutencao THEN
       "RelatorioSAPI".Hora[181] := "SP_Dosagem2";
   END_IF;
   IF "SistemaHabilitado" AND "SinalMisturador1" AND NOT "DosagemContinua_DB3".Manual AND NOT "DosagemContinua_DB3".Manutencao THEN
       "RelatorioSAPI".Hora[182] := "SP_Dosagem3";
   END_IF;
   IF "SistemaHabilitado" AND "SinalMisturador2" AND NOT "DosagemContinua_DB4".Manual AND NOT "DosagemContinua_DB4".Manutencao THEN
       "RelatorioSAPI".Hora[183] := "SP_Dosagem4";
   END_IF;
   IF "SistemaHabilitado" AND "SinalMisturador1" AND NOT "DosagemContinua_DB5".Manual AND NOT "DosagemContinua_DB5".Manutencao THEN
       "RelatorioSAPI".Hora[184] := "SP_Dosagem5";
   END_IF;
   IF "SistemaHabilitado" AND "SinalMisturador2" AND NOT "DosagemContinua_DB6".Manual AND NOT "DosagemContinua_DB6".Manutencao THEN
       "RelatorioSAPI".Hora[185] := "SP_Dosagem6";
   END_IF;
END_REGION
END_ORGANIZATION_BLOCK

ORGANIZATION_BLOCK "05-RedeModbusRTU"   // OB127, LAD, ProgramCycle
{ S7_Optimized_Access := 'TRUE' }
VERSION : 0.1
   VAR_INPUT
      Initial_Call : Bool;
      Remanence : Bool;
   END_VAR
   VAR_TEMP
      desl : Bool;
   END_VAR
   VAR_TEMP   // added for the SCL form of the ladder/FBD networks
      _w1 : Bool;
      _w2 : Bool;
      _w3 : Bool;
      _w4 : Bool;
   END_VAR
BEGIN

REGION Network 1: First scan até modbus ativar
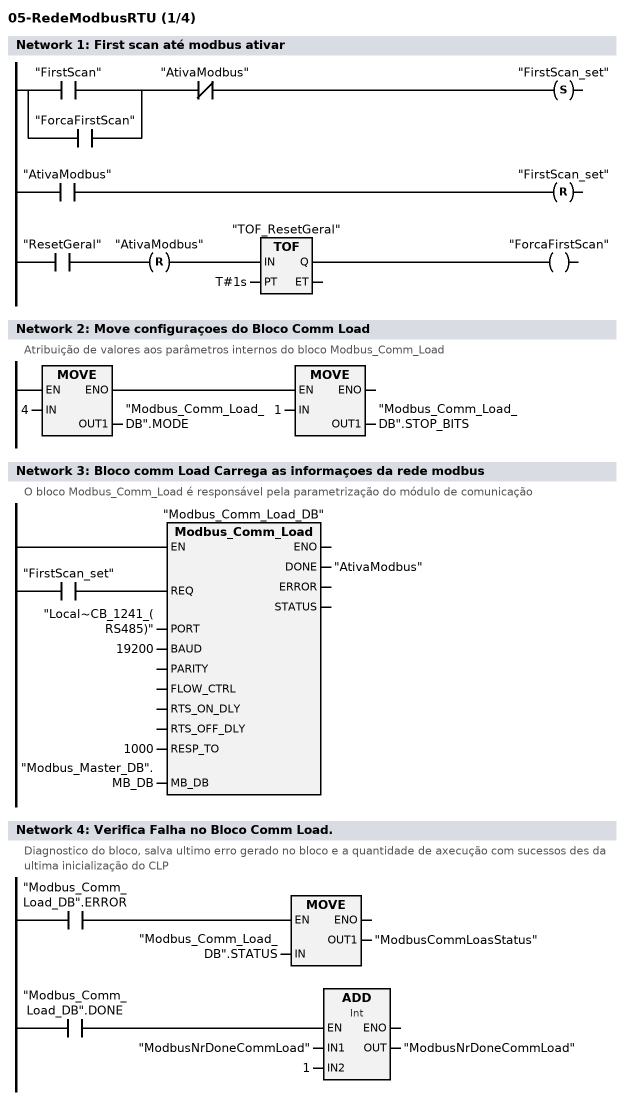
   IF ("FirstScan" OR "ForcaFirstScan") AND NOT "AtivaModbus" THEN "FirstScan_set" := TRUE; END_IF;
   IF "AtivaModbus" THEN "FirstScan_set" := FALSE; END_IF;
   IF "ResetGeral" THEN "AtivaModbus" := FALSE; END_IF;
   "TOF_ResetGeral".TOF(IN := "ResetGeral", PT := T#1s);
   "ForcaFirstScan" := "TOF_ResetGeral".Q;
END_REGION

REGION Network 2: Move configuraçoes do Bloco Comm Load
   // Atribuição de valores aos parâmetros internos do bloco Modbus_Comm_Load
   RUNG wire#powerrail
      Move(in := 4, out1 => "Modbus_Comm_Load_DB".MODE)
      Move(in := 1, out1 => "Modbus_Comm_Load_DB".STOP_BITS)
   END_RUNG
   // the same network as SCL:
   "Modbus_Comm_Load_DB".MODE := 4;
   "Modbus_Comm_Load_DB".STOP_BITS := 1;
END_REGION

REGION Network 3: Bloco comm Load Carrega as informaçoes da rede modbus
   // O bloco Modbus_Comm_Load é responsável pela parametrização do módulo de comunicação
   "Modbus_Comm_Load_DB"(REQ := "FirstScan_set",   // Modbus_Comm_Load
                         PORT := "Local~CB_1241_(RS485)",
                         BAUD := 19200,
                         RESP_TO := 1000,
                         MB_DB := "Modbus_Master_DB".MB_DB,
                         DONE => "AtivaModbus");
END_REGION

REGION Network 4: Verifica Falha no Bloco Comm Load.
   // Diagnostico do bloco, salva ultimo erro gerado no bloco e a quantidade de axecução com sucessos des da ultima inicialização do CLP
   RUNG wire#powerrail
      Contact( "Modbus_Comm_Load_DB".ERROR )
      Move(in := "Modbus_Comm_Load_DB".STATUS, out1 => "ModbusCommLoasStatus")
   END_RUNG
   RUNG wire#powerrail
      Contact( "Modbus_Comm_Load_DB".DONE )
      { S7_Templates := "SrcType := Int" } Add(in1 := "ModbusNrDoneCommLoad", in2 := 1, out => "ModbusNrDoneCommLoad")
   END_RUNG
   // the same network as SCL:
   IF "Modbus_Comm_Load_DB".ERROR THEN "ModbusCommLoasStatus" := "Modbus_Comm_Load_DB".STATUS; END_IF;
   IF "Modbus_Comm_Load_DB".DONE THEN "ModbusNrDoneCommLoad" := "ModbusNrDoneCommLoad" + 1; END_IF;
END_REGION

REGION Network 5: Ponteiro da Rede Modbus
   // Ponteiro da rede de malha fechada, o Index varia entre 1 e 2 e trigger fica em TRUE por um ciclo, após a mudança de estado de Index.
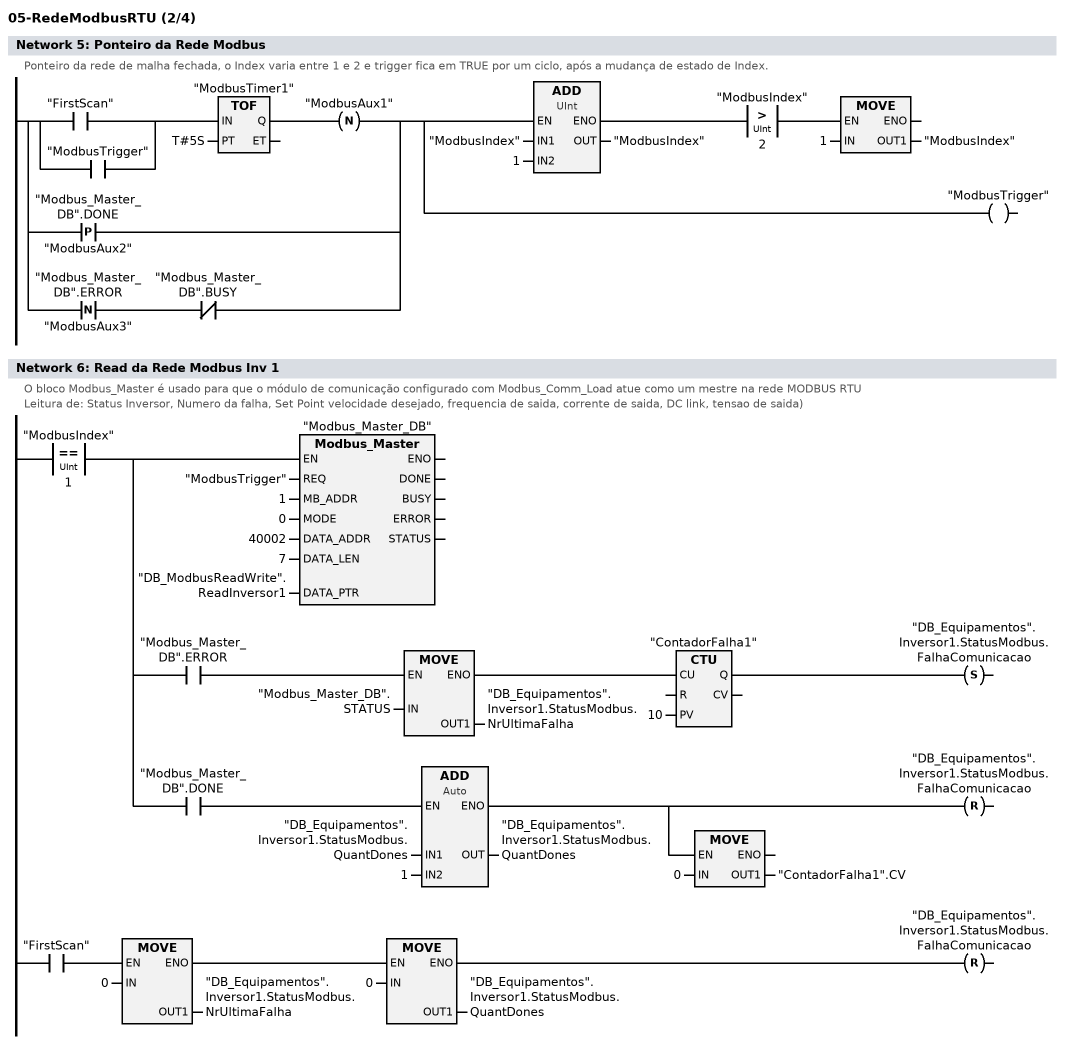
   "ModbusTimer1".TOF(IN := "FirstScan" OR "ModbusTrigger", PT := T#5S);
   #_w1 := NOT "ModbusTimer1".Q AND "ModbusAux1";   // falling edge
   "ModbusAux1" := "ModbusTimer1".Q;
   #_w2 := "Modbus_Master_DB".DONE AND NOT "ModbusAux2";   // rising edge of "Modbus_Master_DB".DONE
   "ModbusAux2" := "Modbus_Master_DB".DONE;
   #_w3 := NOT "Modbus_Master_DB".ERROR AND "ModbusAux3";   // falling edge of "Modbus_Master_DB".ERROR
   "ModbusAux3" := "Modbus_Master_DB".ERROR;
   #_w4 := #_w1 OR #_w2 OR (#_w3 AND NOT "Modbus_Master_DB".BUSY);
   IF #_w4 THEN "ModbusIndex" := "ModbusIndex" + 1; END_IF;
   IF #_w4 AND ("ModbusIndex" > 2) THEN "ModbusIndex" := 1; END_IF;
   "ModbusTrigger" := #_w4;
END_REGION

REGION Network 6: Read da Rede Modbus Inv 1
   // O bloco Modbus_Master é usado para que o módulo de comunicação configurado com Modbus_Comm_Load atue como um mestre na rede MODBUS RTU
   // Leitura de: Status Inversor, Numero da falha, Set Point velocidade desejado, frequencia de saida, corrente de saida, DC link, tensao de saida)
   #_w1 := "ModbusIndex" = 1;
   IF #_w1 THEN
       "Modbus_Master_DB"(REQ := "ModbusTrigger",   // Modbus_Master
                          MB_ADDR := 1,
                          MODE := 0,
                          DATA_ADDR := 40002,
                          DATA_LEN := 7,
                          DATA_PTR := "DB_ModbusReadWrite".ReadInversor1);
   END_IF;
   #_w2 := #_w1 AND "Modbus_Master_DB".ERROR;
   IF #_w2 THEN "DB_Equipamentos".Inversor1.StatusModbus.NrUltimaFalha := "Modbus_Master_DB".STATUS; END_IF;
   "ContadorFalha1".CTU(CU := #_w2, PV := 10);
   IF "ContadorFalha1".Q THEN "DB_Equipamentos".Inversor1.StatusModbus.FalhaComunicacao := TRUE; END_IF;
   IF #_w1 AND "Modbus_Master_DB".DONE THEN
       "DB_Equipamentos".Inversor1.StatusModbus.QuantDones := "DB_Equipamentos".Inversor1.StatusModbus.QuantDones + 1;
       "DB_Equipamentos".Inversor1.StatusModbus.FalhaComunicacao := FALSE;
       "ContadorFalha1".CV := 0;
   END_IF;
   IF "FirstScan" THEN
       "DB_Equipamentos".Inversor1.StatusModbus.NrUltimaFalha := 0;
       "DB_Equipamentos".Inversor1.StatusModbus.QuantDones := 0;
       "DB_Equipamentos".Inversor1.StatusModbus.FalhaComunicacao := FALSE;
   END_IF;
END_REGION

REGION Network 7: Write da Rede Modbus Inv 1
   // O bloco Modbus_Master é usado para que o módulo de comunicação configurado com Modbus_Comm_Load atue como um mestre na rede MODBUS RTU
   // Escrita de valor: CMD e Frequencia
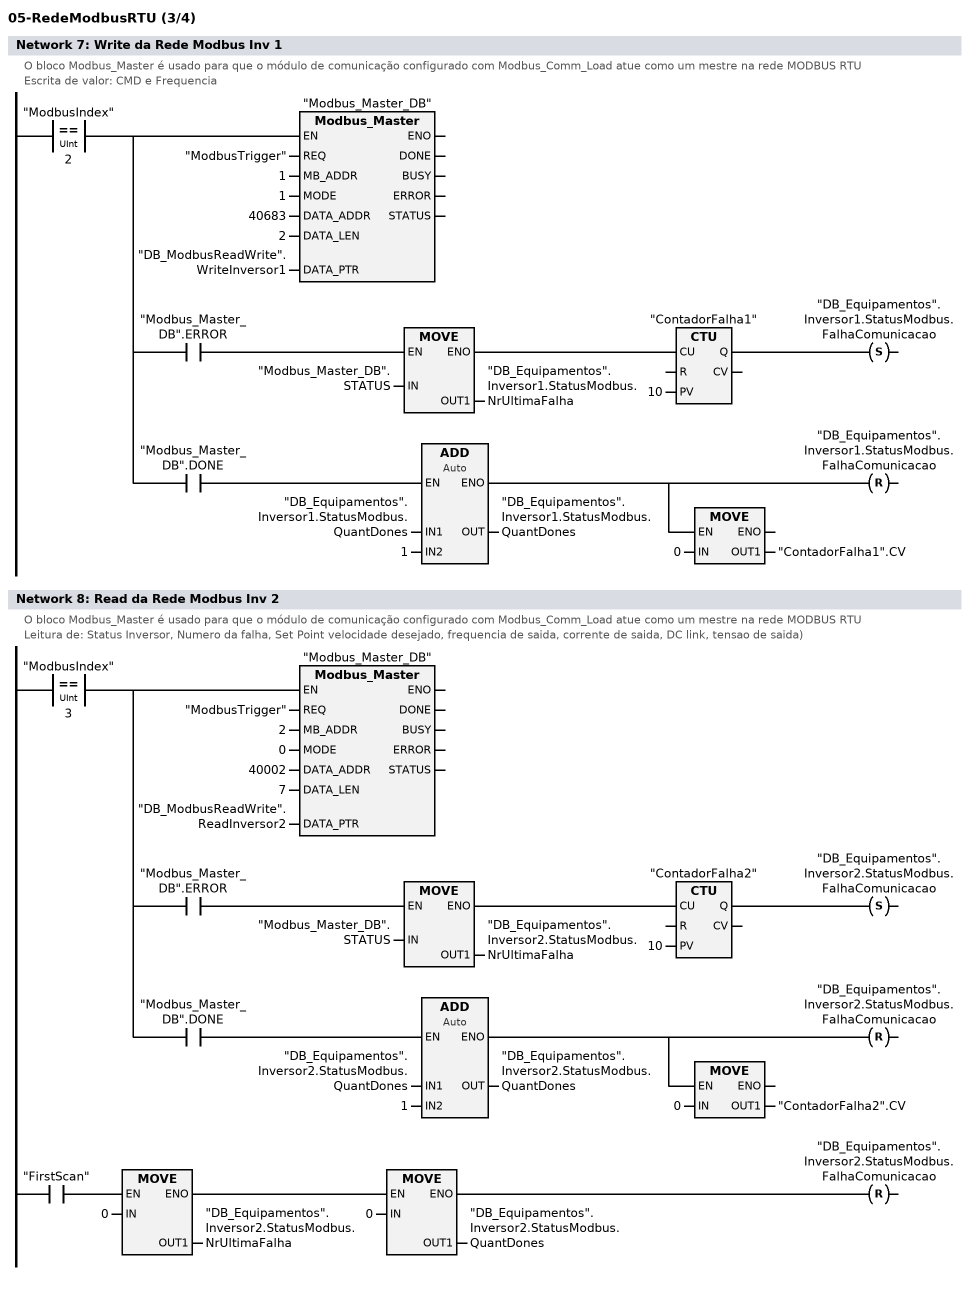
   #_w1 := "ModbusIndex" = 2;
   IF #_w1 THEN
       "Modbus_Master_DB"(REQ := "ModbusTrigger",   // Modbus_Master
                          MB_ADDR := 1,
                          MODE := 1,
                          DATA_ADDR := 40683,
                          DATA_LEN := 2,
                          DATA_PTR := "DB_ModbusReadWrite".WriteInversor1);
   END_IF;
   #_w2 := #_w1 AND "Modbus_Master_DB".ERROR;
   IF #_w2 THEN "DB_Equipamentos".Inversor1.StatusModbus.NrUltimaFalha := "Modbus_Master_DB".STATUS; END_IF;
   "ContadorFalha1".CTU(CU := #_w2, PV := 10);
   IF "ContadorFalha1".Q THEN "DB_Equipamentos".Inversor1.StatusModbus.FalhaComunicacao := TRUE; END_IF;
   IF #_w1 AND "Modbus_Master_DB".DONE THEN
       "DB_Equipamentos".Inversor1.StatusModbus.QuantDones := "DB_Equipamentos".Inversor1.StatusModbus.QuantDones + 1;
       "DB_Equipamentos".Inversor1.StatusModbus.FalhaComunicacao := FALSE;
       "ContadorFalha1".CV := 0;
   END_IF;
END_REGION

REGION Network 8: Read da Rede Modbus Inv 2
   // O bloco Modbus_Master é usado para que o módulo de comunicação configurado com Modbus_Comm_Load atue como um mestre na rede MODBUS RTU
   // Leitura de: Status Inversor, Numero da falha, Set Point velocidade desejado, frequencia de saida, corrente de saida, DC link, tensao de saida)
   #_w1 := "ModbusIndex" = 3;
   IF #_w1 THEN
       "Modbus_Master_DB"(REQ := "ModbusTrigger",   // Modbus_Master
                          MB_ADDR := 2,
                          MODE := 0,
                          DATA_ADDR := 40002,
                          DATA_LEN := 7,
                          DATA_PTR := "DB_ModbusReadWrite".ReadInversor2);
   END_IF;
   #_w2 := #_w1 AND "Modbus_Master_DB".ERROR;
   IF #_w2 THEN "DB_Equipamentos".Inversor2.StatusModbus.NrUltimaFalha := "Modbus_Master_DB".STATUS; END_IF;
   "ContadorFalha2".CTU(CU := #_w2, PV := 10);
   IF "ContadorFalha2".Q THEN "DB_Equipamentos".Inversor2.StatusModbus.FalhaComunicacao := TRUE; END_IF;
   IF #_w1 AND "Modbus_Master_DB".DONE THEN
       "DB_Equipamentos".Inversor2.StatusModbus.QuantDones := "DB_Equipamentos".Inversor2.StatusModbus.QuantDones + 1;
       "DB_Equipamentos".Inversor2.StatusModbus.FalhaComunicacao := FALSE;
       "ContadorFalha2".CV := 0;
   END_IF;
   IF "FirstScan" THEN
       "DB_Equipamentos".Inversor2.StatusModbus.NrUltimaFalha := 0;
       "DB_Equipamentos".Inversor2.StatusModbus.QuantDones := 0;
       "DB_Equipamentos".Inversor2.StatusModbus.FalhaComunicacao := FALSE;
   END_IF;
END_REGION

REGION Network 9: Write da Rede Modbus Inv 2
   // O bloco Modbus_Master é usado para que o módulo de comunicação configurado com Modbus_Comm_Load atue como um mestre na rede MODBUS RTU
   // Escrita de valor: CMD e Frequencia
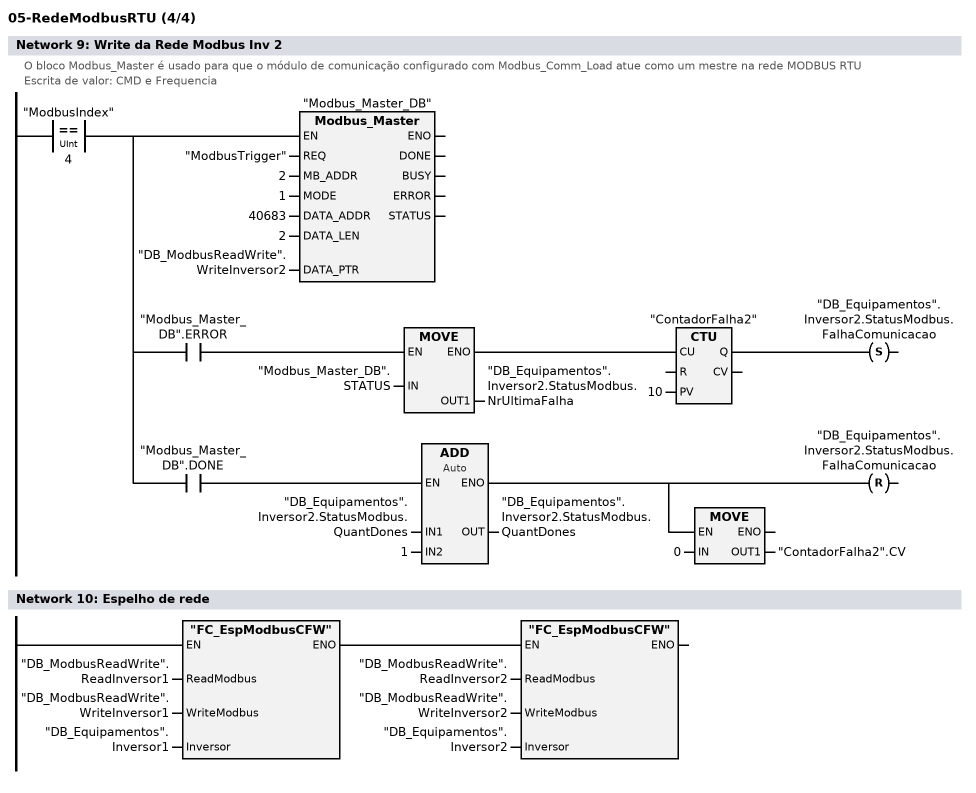
   #_w1 := "ModbusIndex" = 4;
   IF #_w1 THEN
       "Modbus_Master_DB"(REQ := "ModbusTrigger",   // Modbus_Master
                          MB_ADDR := 2,
                          MODE := 1,
                          DATA_ADDR := 40683,
                          DATA_LEN := 2,
                          DATA_PTR := "DB_ModbusReadWrite".WriteInversor2);
   END_IF;
   #_w2 := #_w1 AND "Modbus_Master_DB".ERROR;
   IF #_w2 THEN "DB_Equipamentos".Inversor2.StatusModbus.NrUltimaFalha := "Modbus_Master_DB".STATUS; END_IF;
   "ContadorFalha2".CTU(CU := #_w2, PV := 10);
   IF "ContadorFalha2".Q THEN "DB_Equipamentos".Inversor2.StatusModbus.FalhaComunicacao := TRUE; END_IF;
   IF #_w1 AND "Modbus_Master_DB".DONE THEN
       "DB_Equipamentos".Inversor2.StatusModbus.QuantDones := "DB_Equipamentos".Inversor2.StatusModbus.QuantDones + 1;
       "DB_Equipamentos".Inversor2.StatusModbus.FalhaComunicacao := FALSE;
       "ContadorFalha2".CV := 0;
   END_IF;
END_REGION

REGION Network 10: Espelho de rede
   RUNG wire#powerrail
      "FC_EspModbusCFW"(ReadModbus := "DB_ModbusReadWrite".ReadInversor1, WriteModbus := "DB_ModbusReadWrite".WriteInversor1, Inversor := "DB_Equipamentos".Inversor1)
      "FC_EspModbusCFW"(ReadModbus := "DB_ModbusReadWrite".ReadInversor2, WriteModbus := "DB_ModbusReadWrite".WriteInversor2, Inversor := "DB_Equipamentos".Inversor2)
   END_RUNG
   // the same network as SCL:
   "FC_EspModbusCFW"(ReadModbus := "DB_ModbusReadWrite".ReadInversor1,
                     WriteModbus := "DB_ModbusReadWrite".WriteInversor1,
                     Inversor := "DB_Equipamentos".Inversor1,
                     ENO => #_w1);
   IF #_w1 THEN
       "FC_EspModbusCFW"(ReadModbus := "DB_ModbusReadWrite".ReadInversor2,
                         WriteModbus := "DB_ModbusReadWrite".WriteInversor2,
                         Inversor := "DB_Equipamentos".Inversor2);
   END_IF;
END_REGION
END_ORGANIZATION_BLOCK

ORGANIZATION_BLOCK "06-Integracao"   // OB128, LAD, ProgramCycle
{ S7_Optimized_Access := 'TRUE' }
VERSION : 0.1
   VAR_INPUT
      Initial_Call : Bool;
      Remanence : Bool;
   END_VAR
   VAR_TEMP   // added for the SCL form of the ladder/FBD networks
      _w1 : Bool;
   END_VAR
BEGIN

REGION Network 1: Put e falha de comunicação
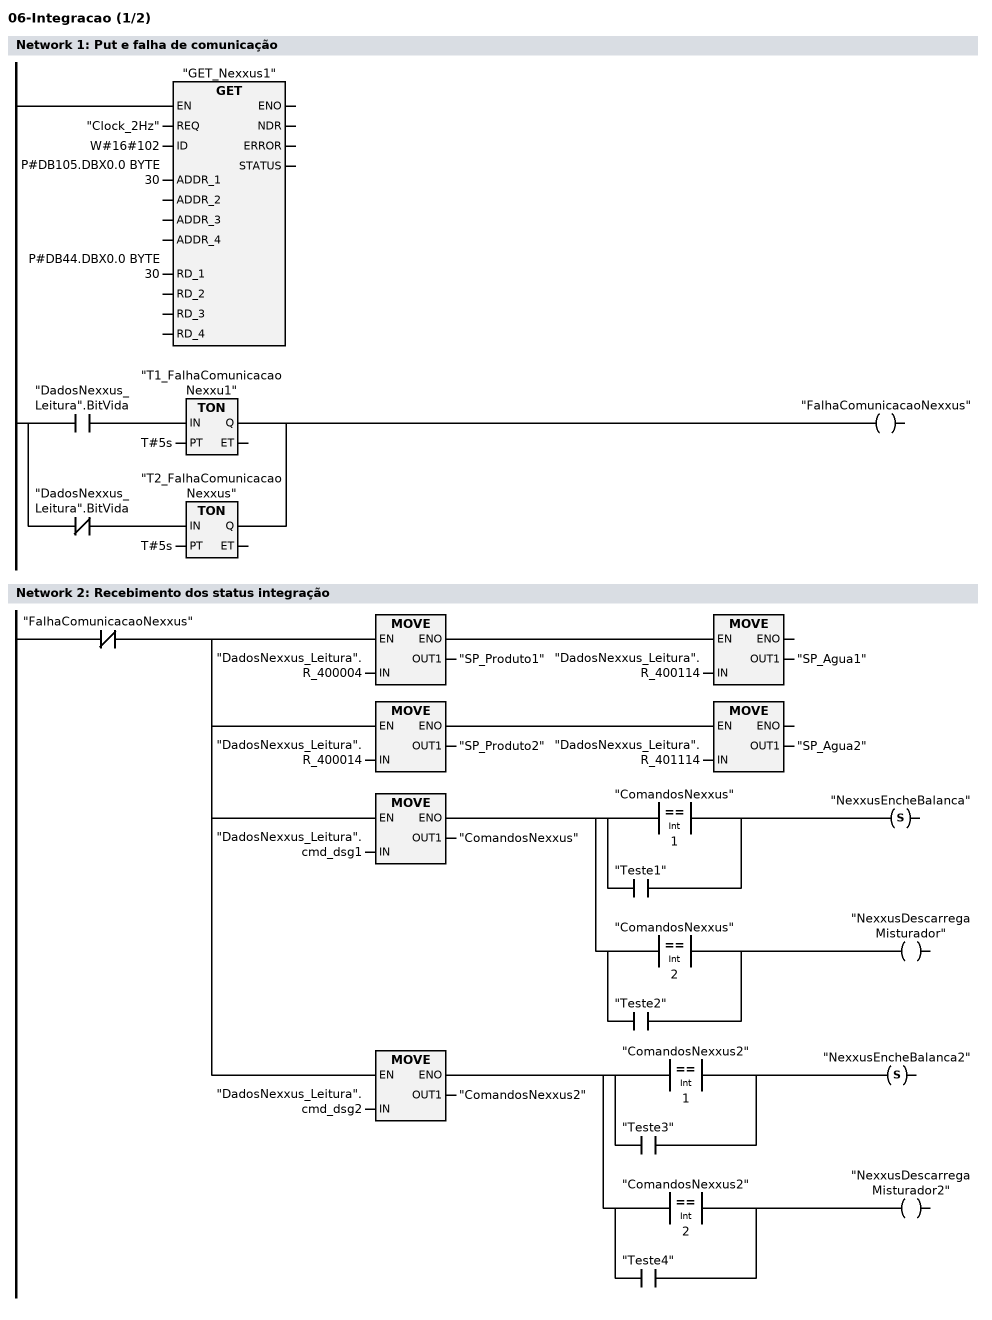
   "GET_Nexxus1"(REQ := "Clock_2Hz",   // GET
                 ID := W#16#102,
                 ADDR_1 := P#DB105.DBX0.0 BYTE 30,
                 RD_1 := P#DB44.DBX0.0 BYTE 30);
   "T1_FalhaComunicacaoNexxu1".TON(IN := "DadosNexxus_Leitura".BitVida, PT := T#5s);
   "T2_FalhaComunicacaoNexxus".TON(IN := NOT "DadosNexxus_Leitura".BitVida, PT := T#5s);
   "FalhaComunicacaoNexxus" := "T1_FalhaComunicacaoNexxu1".Q OR "T2_FalhaComunicacaoNexxus".Q;
END_REGION

REGION Network 2: Recebimento dos status integração
   RUNG wire#powerrail
      I_Contact( "FalhaComunicacaoNexxus" )
      wire#w1
      Move(in := "DadosNexxus_Leitura".R_400004, out1 => "SP_Produto1")
      Move(in := "DadosNexxus_Leitura".R_400114, out1 => "SP_Agua1")
   END_RUNG
   RUNG wire#w1
      Move(in := "DadosNexxus_Leitura".R_400014, out1 => "SP_Produto2")
      Move(in := "DadosNexxus_Leitura".R_401114, out1 => "SP_Agua2")
   END_RUNG
   RUNG wire#w1
      Move(in := "DadosNexxus_Leitura".cmd_dsg1, out1 => "ComandosNexxus")
      wire#w2
      { S7_Templates := "SrcType := Int" } EQ_Contact(in1 := "ComandosNexxus", in2 := 1)
      wire#w3
      S_Coil( "NexxusEncheBalanca" )
   END_RUNG
   RUNG wire#w2
      Contact( "Teste1" )
   END_RUNG wire#w3
   RUNG wire#w2
      { S7_Templates := "SrcType := Int" } EQ_Contact(in1 := "ComandosNexxus", in2 := 2)
      wire#w4
      Coil( "NexxusDescarregaMisturador" )
   END_RUNG
   RUNG wire#w2
      Contact( "Teste2" )
   END_RUNG wire#w4
   RUNG wire#w1
      Move(in := "DadosNexxus_Leitura".cmd_dsg2, out1 => "ComandosNexxus2")
      wire#w5
      { S7_Templates := "SrcType := Int" } EQ_Contact(in1 := "ComandosNexxus2", in2 := 1)
      wire#w6
      S_Coil( "NexxusEncheBalanca2" )
   END_RUNG
   RUNG wire#w5
      Contact( "Teste3" )
   END_RUNG wire#w6
   RUNG wire#w5
      { S7_Templates := "SrcType := Int" } EQ_Contact(in1 := "ComandosNexxus2", in2 := 2)
      wire#w7
      Coil( "NexxusDescarregaMisturador2" )
   END_RUNG
   RUNG wire#w5
      Contact( "Teste4" )
   END_RUNG wire#w7
   // the same network as SCL:
   #_w1 := NOT "FalhaComunicacaoNexxus";
   IF #_w1 THEN
       "SP_Produto1" := "DadosNexxus_Leitura".R_400004;
       "SP_Agua1" := "DadosNexxus_Leitura".R_400114;
       "SP_Produto2" := "DadosNexxus_Leitura".R_400014;
       "SP_Agua2" := "DadosNexxus_Leitura".R_401114;
       "ComandosNexxus" := "DadosNexxus_Leitura".cmd_dsg1;
   END_IF;
   IF #_w1 AND (("ComandosNexxus" = 1) OR "Teste1") THEN "NexxusEncheBalanca" := TRUE; END_IF;
   "NexxusDescarregaMisturador" := #_w1 AND (("ComandosNexxus" = 2) OR "Teste2");
   IF #_w1 THEN "ComandosNexxus2" := "DadosNexxus_Leitura".cmd_dsg2; END_IF;
   IF #_w1 AND (("ComandosNexxus2" = 1) OR "Teste3") THEN "NexxusEncheBalanca2" := TRUE; END_IF;
   "NexxusDescarregaMisturador2" := #_w1 AND (("ComandosNexxus2" = 2) OR "Teste4");
END_REGION

REGION Network 3: Escrita para Nexxus
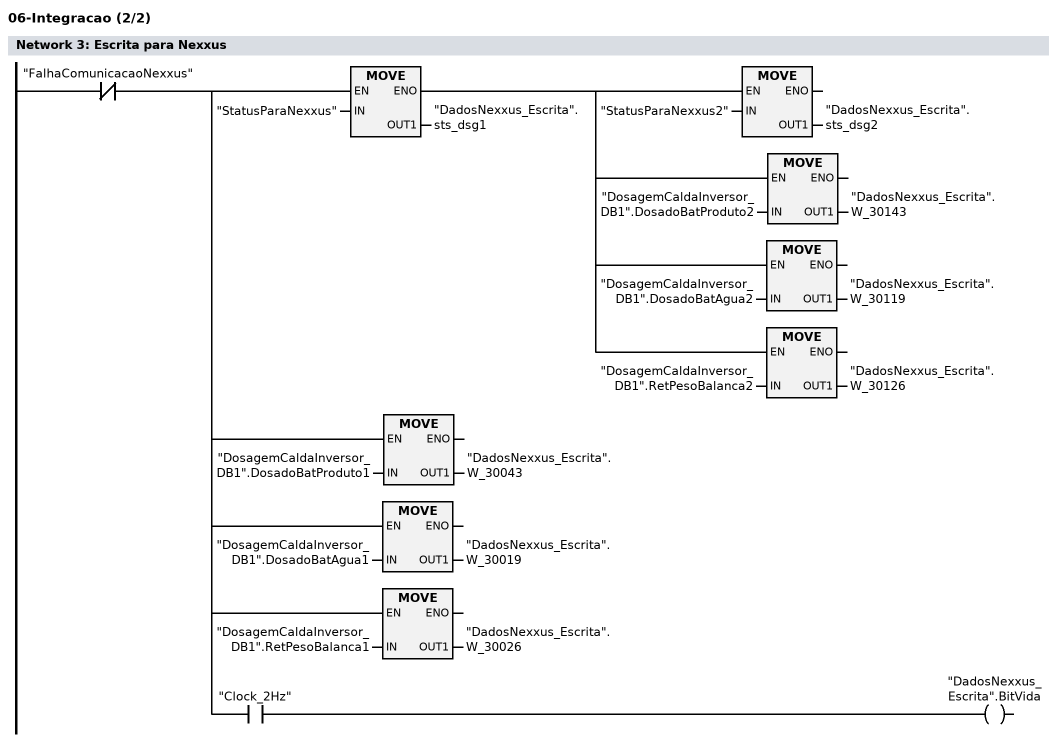
   RUNG wire#powerrail
      I_Contact( "FalhaComunicacaoNexxus" )
      wire#w1
      Move(in := "StatusParaNexxus", out1 => "DadosNexxus_Escrita".sts_dsg1)
      wire#w2
      Move(in := "StatusParaNexxus2", out1 => "DadosNexxus_Escrita".sts_dsg2)
   END_RUNG
   RUNG wire#w2
      Move(in := "DosagemCaldaInversor_DB1".DosadoBatProduto2, out1 => "DadosNexxus_Escrita".W_30143)
   END_RUNG
   RUNG wire#w2
      Move(in := "DosagemCaldaInversor_DB1".DosadoBatAgua2, out1 => "DadosNexxus_Escrita".W_30119)
   END_RUNG
   RUNG wire#w2
      Move(in := "DosagemCaldaInversor_DB1".RetPesoBalanca2, out1 => "DadosNexxus_Escrita".W_30126)
   END_RUNG
   RUNG wire#w1
      Move(in := "DosagemCaldaInversor_DB1".DosadoBatProduto1, out1 => "DadosNexxus_Escrita".W_30043)
   END_RUNG
   RUNG wire#w1
      Move(in := "DosagemCaldaInversor_DB1".DosadoBatAgua1, out1 => "DadosNexxus_Escrita".W_30019)
   END_RUNG
   RUNG wire#w1
      Move(in := "DosagemCaldaInversor_DB1".RetPesoBalanca1, out1 => "DadosNexxus_Escrita".W_30026)
   END_RUNG
   RUNG wire#w1
      Contact( "Clock_2Hz" )
      Coil( "DadosNexxus_Escrita".BitVida )
   END_RUNG
   // the same network as SCL:
   #_w1 := NOT "FalhaComunicacaoNexxus";
   IF #_w1 THEN
       "DadosNexxus_Escrita".sts_dsg1 := "StatusParaNexxus";
       "DadosNexxus_Escrita".sts_dsg2 := "StatusParaNexxus2";
       "DadosNexxus_Escrita".W_30143 := "DosagemCaldaInversor_DB1".DosadoBatProduto2;
       "DadosNexxus_Escrita".W_30119 := "DosagemCaldaInversor_DB1".DosadoBatAgua2;
       "DadosNexxus_Escrita".W_30126 := "DosagemCaldaInversor_DB1".RetPesoBalanca2;
       "DadosNexxus_Escrita".W_30043 := "DosagemCaldaInversor_DB1".DosadoBatProduto1;
       "DadosNexxus_Escrita".W_30019 := "DosagemCaldaInversor_DB1".DosadoBatAgua1;
       "DadosNexxus_Escrita".W_30026 := "DosagemCaldaInversor_DB1".RetPesoBalanca1;
   END_IF;
   "DadosNexxus_Escrita".BitVida := #_w1 AND "Clock_2Hz";
END_REGION
END_ORGANIZATION_BLOCK

// folder: FB

FUNCTION_BLOCK "InputClp"   // FB1, LAD
{ S7_Optimized_Access := 'TRUE' }
VERSION : 0.1
   VAR_INPUT
      "DI.a.0" : Bool;
      "DI.a.1" : Bool;
      "DI.a.2" : Bool;
      "DI.a.3" : Bool;
      "DI.a.4" : Bool;
      "DI.a.5" : Bool;
      "DI.a.6" : Bool;
      "DI.a.7" : Bool;
      "DI.b.0" : Bool;
      "DI.b.1" : Bool;
      "DI.b.2" : Bool;
      "DI.b.3" : Bool;
      "DI.b.4" : Bool;
      "DI.b.5" : Bool;
   END_VAR
   VAR_OUTPUT
      "DI.0.0" : Bool;
      "DI.0.1" : Bool;
      "DI.0.2" : Bool;
      "DI.0.3" : Bool;
      "DI.0.4" : Bool;
      "DI.0.5" : Bool;
      "DI.0.6" : Bool;
      "DI.0.7" : Bool;
      "DI.1.0" : Bool;
      "DI.1.1" : Bool;
      "DI.1.2" : Bool;
      "DI.1.3" : Bool;
      "DI.1.4" : Bool;
      "DI.1.5" : Bool;
   END_VAR
   VAR
      ForcaDIa0 : Bool;
      ForcaDIa1 : Bool;
      ForcaDIa2 : Bool;
      ForcaDIa3 : Bool;
      ForcaDIa4 : Bool;
      ForcaDIa5 : Bool;
      ForcaDIa6 : Bool;
      ForcaDIa7 : Bool;
      ForcaDIb0 : Bool;
      ForcaDIb1 : Bool;
      ForcaDIb2 : Bool;
      ForcaDIb3 : Bool;
      ForcaDIb4 : Bool;
      ForcaDIb5 : Bool;
   END_VAR
BEGIN

REGION Network 1
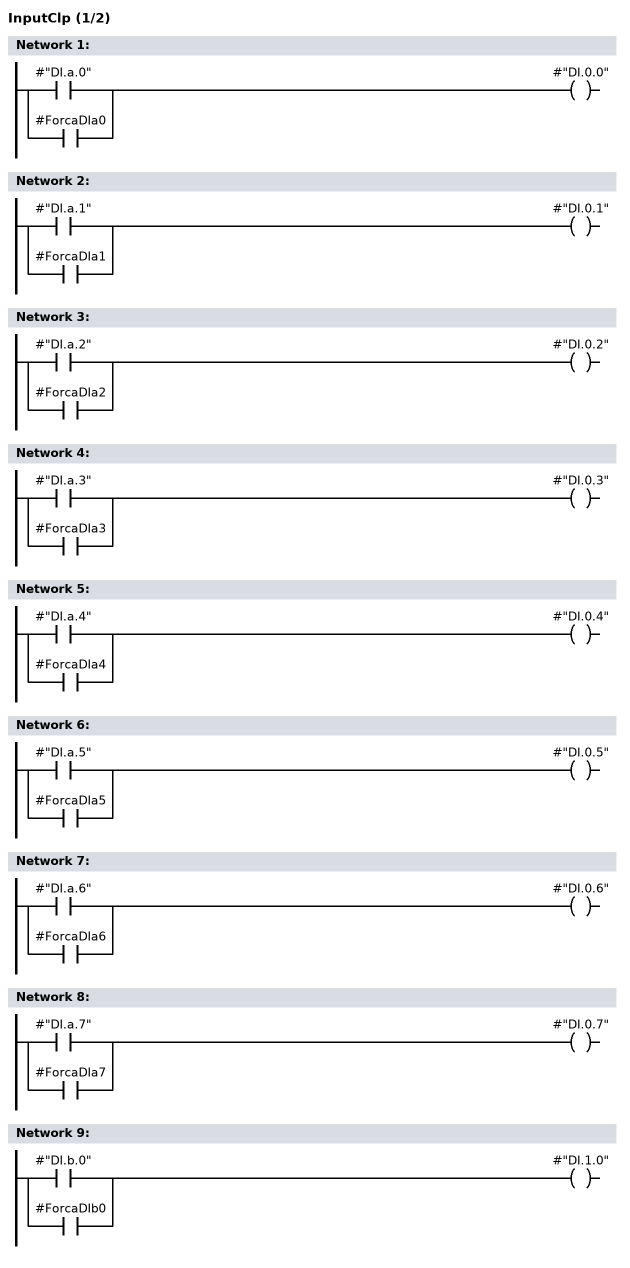
   RUNG wire#powerrail
      Contact( #"DI.a.0" )
      wire#w1
      Coil( #"DI.0.0" )
   END_RUNG
   RUNG wire#powerrail
      Contact( #ForcaDIa0 )
   END_RUNG wire#w1
   // the same network as SCL:
   #"DI.0.0" := #"DI.a.0" OR #ForcaDIa0;
END_REGION

REGION Network 2
   RUNG wire#powerrail
      Contact( #"DI.a.1" )
      wire#w1
      Coil( #"DI.0.1" )
   END_RUNG
   RUNG wire#powerrail
      Contact( #ForcaDIa1 )
   END_RUNG wire#w1
   // the same network as SCL:
   #"DI.0.1" := #"DI.a.1" OR #ForcaDIa1;
END_REGION

REGION Network 3
   RUNG wire#powerrail
      Contact( #"DI.a.2" )
      wire#w1
      Coil( #"DI.0.2" )
   END_RUNG
   RUNG wire#powerrail
      Contact( #ForcaDIa2 )
   END_RUNG wire#w1
   // the same network as SCL:
   #"DI.0.2" := #"DI.a.2" OR #ForcaDIa2;
END_REGION

REGION Network 4
   RUNG wire#powerrail
      Contact( #"DI.a.3" )
      wire#w1
      Coil( #"DI.0.3" )
   END_RUNG
   RUNG wire#powerrail
      Contact( #ForcaDIa3 )
   END_RUNG wire#w1
   // the same network as SCL:
   #"DI.0.3" := #"DI.a.3" OR #ForcaDIa3;
END_REGION

REGION Network 5
   RUNG wire#powerrail
      Contact( #"DI.a.4" )
      wire#w1
      Coil( #"DI.0.4" )
   END_RUNG
   RUNG wire#powerrail
      Contact( #ForcaDIa4 )
   END_RUNG wire#w1
   // the same network as SCL:
   #"DI.0.4" := #"DI.a.4" OR #ForcaDIa4;
END_REGION

REGION Network 6
   RUNG wire#powerrail
      Contact( #"DI.a.5" )
      wire#w1
      Coil( #"DI.0.5" )
   END_RUNG
   RUNG wire#powerrail
      Contact( #ForcaDIa5 )
   END_RUNG wire#w1
   // the same network as SCL:
   #"DI.0.5" := #"DI.a.5" OR #ForcaDIa5;
END_REGION

REGION Network 7
   RUNG wire#powerrail
      Contact( #"DI.a.6" )
      wire#w1
      Coil( #"DI.0.6" )
   END_RUNG
   RUNG wire#powerrail
      Contact( #ForcaDIa6 )
   END_RUNG wire#w1
   // the same network as SCL:
   #"DI.0.6" := #"DI.a.6" OR #ForcaDIa6;
END_REGION

REGION Network 8
   RUNG wire#powerrail
      Contact( #"DI.a.7" )
      wire#w1
      Coil( #"DI.0.7" )
   END_RUNG
   RUNG wire#powerrail
      Contact( #ForcaDIa7 )
   END_RUNG wire#w1
   // the same network as SCL:
   #"DI.0.7" := #"DI.a.7" OR #ForcaDIa7;
END_REGION

REGION Network 9
   RUNG wire#powerrail
      Contact( #"DI.b.0" )
      wire#w1
      Coil( #"DI.1.0" )
   END_RUNG
   RUNG wire#powerrail
      Contact( #ForcaDIb0 )
   END_RUNG wire#w1
   // the same network as SCL:
   #"DI.1.0" := #"DI.b.0" OR #ForcaDIb0;
END_REGION

REGION Network 10
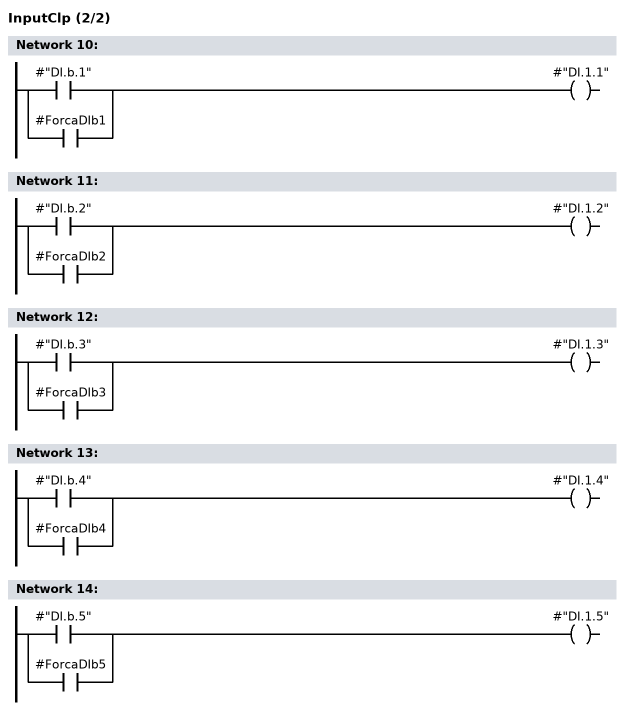
   RUNG wire#powerrail
      Contact( #"DI.b.1" )
      wire#w1
      Coil( #"DI.1.1" )
   END_RUNG
   RUNG wire#powerrail
      Contact( #ForcaDIb1 )
   END_RUNG wire#w1
   // the same network as SCL:
   #"DI.1.1" := #"DI.b.1" OR #ForcaDIb1;
END_REGION

REGION Network 11
   RUNG wire#powerrail
      Contact( #"DI.b.2" )
      wire#w1
      Coil( #"DI.1.2" )
   END_RUNG
   RUNG wire#powerrail
      Contact( #ForcaDIb2 )
   END_RUNG wire#w1
   // the same network as SCL:
   #"DI.1.2" := #"DI.b.2" OR #ForcaDIb2;
END_REGION

REGION Network 12
   RUNG wire#powerrail
      Contact( #"DI.b.3" )
      wire#w1
      Coil( #"DI.1.3" )
   END_RUNG
   RUNG wire#powerrail
      Contact( #ForcaDIb3 )
   END_RUNG wire#w1
   // the same network as SCL:
   #"DI.1.3" := #"DI.b.3" OR #ForcaDIb3;
END_REGION

REGION Network 13
   RUNG wire#powerrail
      Contact( #"DI.b.4" )
      wire#w1
      Coil( #"DI.1.4" )
   END_RUNG
   RUNG wire#powerrail
      Contact( #ForcaDIb4 )
   END_RUNG wire#w1
   // the same network as SCL:
   #"DI.1.4" := #"DI.b.4" OR #ForcaDIb4;
END_REGION

REGION Network 14
   RUNG wire#powerrail
      Contact( #"DI.b.5" )
      wire#w1
      Coil( #"DI.1.5" )
   END_RUNG
   RUNG wire#powerrail
      Contact( #ForcaDIb5 )
   END_RUNG wire#w1
   // the same network as SCL:
   #"DI.1.5" := #"DI.b.5" OR #ForcaDIb5;
END_REGION
END_FUNCTION_BLOCK

FUNCTION_BLOCK "OutputClp"   // FB2, LAD
{ S7_Optimized_Access := 'TRUE' }
VERSION : 0.1
   VAR_INPUT
      "DO.a.0" : Bool;
      "DO.a.1" : Bool;
      "DO.a.2" : Bool;
      "DO.a.3" : Bool;
      "DO.a.4" : Bool;
      "DO.a.5" : Bool;
      "DO.a.6" : Bool;
      "DO.a.7" : Bool;
      "DO.b.0" : Bool;
      "DO.b.1" : Bool;
   END_VAR
   VAR_OUTPUT
      "DO.0.0" : Bool;
      "DO.0.1" : Bool;
      "DO.0.2" : Bool;
      "DO.0.3" : Bool;
      "DO.0.4" : Bool;
      "DO.0.5" : Bool;
      "DO.0.6" : Bool;
      "DO.0.7" : Bool;
      "DO.1.0" : Bool;
      "DO.1.1" : Bool;
   END_VAR
   VAR
      ForcaDOa0 : Bool;
      ForcaDOa1 : Bool;
      ForcaDOa2 : Bool;
      ForcaDOa3 : Bool;
      ForcaDOa4 : Bool;
      ForcaDOa5 : Bool;
      ForcaDOa6 : Bool;
      ForcaDOa7 : Bool;
      ForcaDOb0 : Bool;
      ForcaDOb1 : Bool;
   END_VAR
BEGIN

REGION Network 1
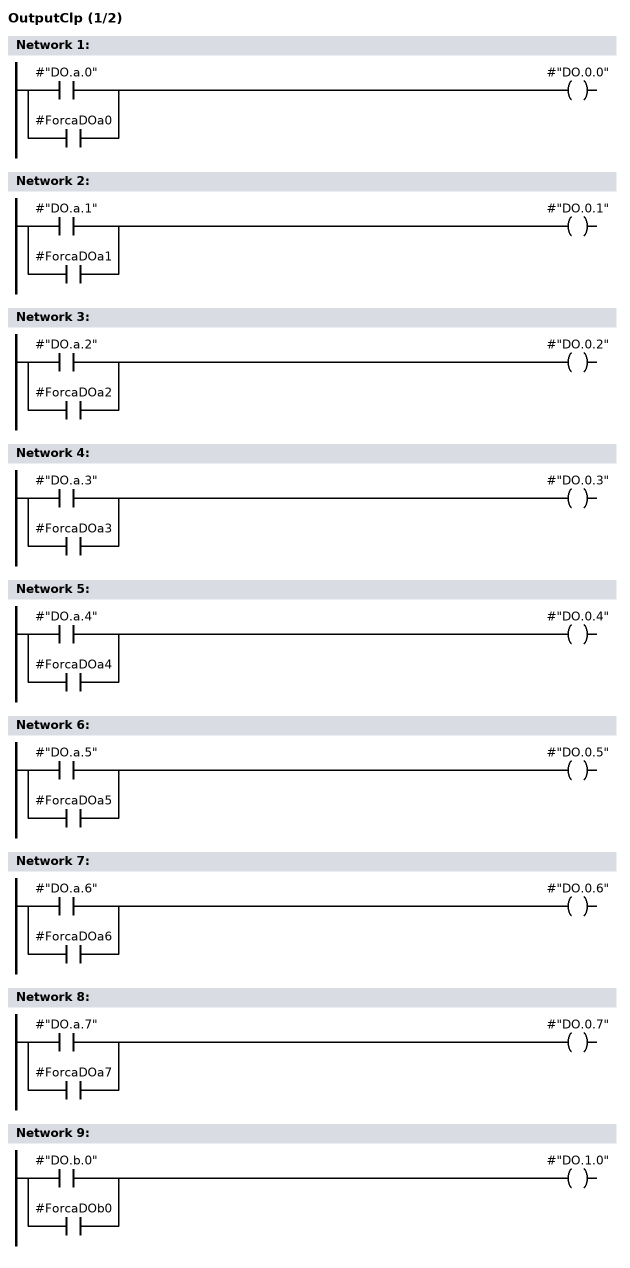
   RUNG wire#powerrail
      Contact( #"DO.a.0" )
      wire#w1
      Coil( #"DO.0.0" )
   END_RUNG
   RUNG wire#powerrail
      Contact( #ForcaDOa0 )
   END_RUNG wire#w1
   // the same network as SCL:
   #"DO.0.0" := #"DO.a.0" OR #ForcaDOa0;
END_REGION

REGION Network 2
   RUNG wire#powerrail
      Contact( #"DO.a.1" )
      wire#w1
      Coil( #"DO.0.1" )
   END_RUNG
   RUNG wire#powerrail
      Contact( #ForcaDOa1 )
   END_RUNG wire#w1
   // the same network as SCL:
   #"DO.0.1" := #"DO.a.1" OR #ForcaDOa1;
END_REGION

REGION Network 3
   RUNG wire#powerrail
      Contact( #"DO.a.2" )
      wire#w1
      Coil( #"DO.0.2" )
   END_RUNG
   RUNG wire#powerrail
      Contact( #ForcaDOa2 )
   END_RUNG wire#w1
   // the same network as SCL:
   #"DO.0.2" := #"DO.a.2" OR #ForcaDOa2;
END_REGION

REGION Network 4
   RUNG wire#powerrail
      Contact( #"DO.a.3" )
      wire#w1
      Coil( #"DO.0.3" )
   END_RUNG
   RUNG wire#powerrail
      Contact( #ForcaDOa3 )
   END_RUNG wire#w1
   // the same network as SCL:
   #"DO.0.3" := #"DO.a.3" OR #ForcaDOa3;
END_REGION

REGION Network 5
   RUNG wire#powerrail
      Contact( #"DO.a.4" )
      wire#w1
      Coil( #"DO.0.4" )
   END_RUNG
   RUNG wire#powerrail
      Contact( #ForcaDOa4 )
   END_RUNG wire#w1
   // the same network as SCL:
   #"DO.0.4" := #"DO.a.4" OR #ForcaDOa4;
END_REGION

REGION Network 6
   RUNG wire#powerrail
      Contact( #"DO.a.5" )
      wire#w1
      Coil( #"DO.0.5" )
   END_RUNG
   RUNG wire#powerrail
      Contact( #ForcaDOa5 )
   END_RUNG wire#w1
   // the same network as SCL:
   #"DO.0.5" := #"DO.a.5" OR #ForcaDOa5;
END_REGION

REGION Network 7
   RUNG wire#powerrail
      Contact( #"DO.a.6" )
      wire#w1
      Coil( #"DO.0.6" )
   END_RUNG
   RUNG wire#powerrail
      Contact( #ForcaDOa6 )
   END_RUNG wire#w1
   // the same network as SCL:
   #"DO.0.6" := #"DO.a.6" OR #ForcaDOa6;
END_REGION

REGION Network 8
   RUNG wire#powerrail
      Contact( #"DO.a.7" )
      wire#w1
      Coil( #"DO.0.7" )
   END_RUNG
   RUNG wire#powerrail
      Contact( #ForcaDOa7 )
   END_RUNG wire#w1
   // the same network as SCL:
   #"DO.0.7" := #"DO.a.7" OR #ForcaDOa7;
END_REGION

REGION Network 9
   RUNG wire#powerrail
      Contact( #"DO.b.0" )
      wire#w1
      Coil( #"DO.1.0" )
   END_RUNG
   RUNG wire#powerrail
      Contact( #ForcaDOb0 )
   END_RUNG wire#w1
   // the same network as SCL:
   #"DO.1.0" := #"DO.b.0" OR #ForcaDOb0;
END_REGION

REGION Network 10
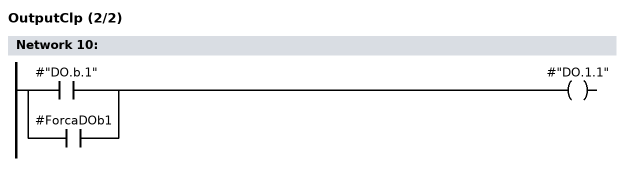
   RUNG wire#powerrail
      Contact( #"DO.b.1" )
      wire#w1
      Coil( #"DO.1.1" )
   END_RUNG
   RUNG wire#powerrail
      Contact( #ForcaDOb1 )
   END_RUNG wire#w1
   // the same network as SCL:
   #"DO.1.1" := #"DO.b.1" OR #ForcaDOb1;
END_REGION
END_FUNCTION_BLOCK

FUNCTION_BLOCK "InputMod16"   // FB3, LAD
{ S7_Optimized_Access := 'TRUE' }
VERSION : 0.1
   VAR_INPUT
      "DI.a.0" : Bool;
      "DI.a.1" : Bool;
      "DI.a.2" : Bool;
      "DI.a.3" : Bool;
      "DI.a.4" : Bool;
      "DI.a.5" : Bool;
      "DI.a.6" : Bool;
      "DI.a.7" : Bool;
      "DI.b.0" : Bool;
      "DI.b.1" : Bool;
      "DI.b.2" : Bool;
      "DI.b.3" : Bool;
      "DI.b.4" : Bool;
      "DI.b.5" : Bool;
      "DI.b.6" : Bool;
      "DI.b.7" : Bool;
   END_VAR
   VAR_OUTPUT
      "DI.0.0" : Bool;
      "DI.0.1" : Bool;
      "DI.0.2" : Bool;
      "DI.0.3" : Bool;
      "DI.0.4" : Bool;
      "DI.0.5" : Bool;
      "DI.0.6" : Bool;
      "DI.0.7" : Bool;
      "DI.1.0" : Bool;
      "DI.1.1" : Bool;
      "DI.1.2" : Bool;
      "DI.1.3" : Bool;
      "DI.1.4" : Bool;
      "DI.1.5" : Bool;
      "DI.1.6" : Bool;
      "DI.1.7" : Bool;
   END_VAR
   VAR
      ForcaDIa0 : Bool;
      ForcaDIa1 : Bool;
      ForcaDIa2 : Bool;
      ForcaDIa3 : Bool;
      ForcaDIa4 : Bool;
      ForcaDIa5 : Bool;
      ForcaDIa6 : Bool;
      ForcaDIa7 : Bool;
      ForcaDIb0 : Bool;
      ForcaDIb1 : Bool;
      ForcaDIb2 : Bool;
      ForcaDIb3 : Bool;
      ForcaDIb4 : Bool;
      ForcaDIb5 : Bool;
      ForcaDIb6 : Bool;
      ForcaDIb7 : Bool;
   END_VAR
BEGIN

REGION Network 1
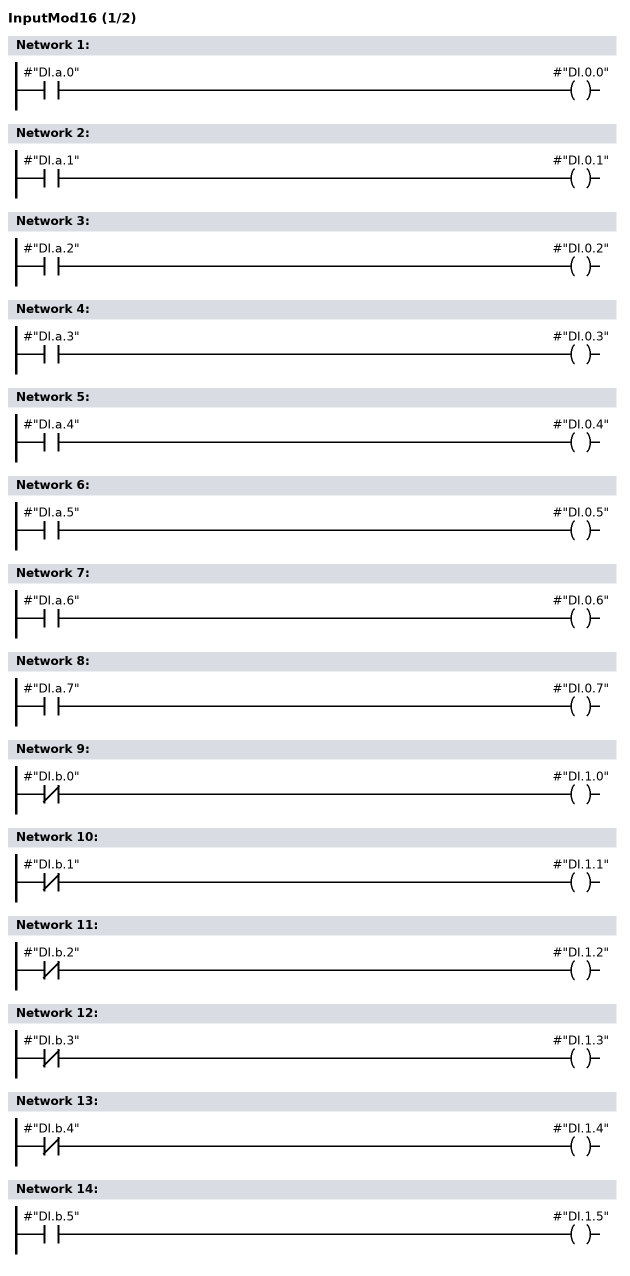
   RUNG wire#powerrail
      Contact( #"DI.a.0" )
      Coil( #"DI.0.0" )
   END_RUNG
   // the same network as SCL:
   #"DI.0.0" := #"DI.a.0";
END_REGION

REGION Network 2
   RUNG wire#powerrail
      Contact( #"DI.a.1" )
      Coil( #"DI.0.1" )
   END_RUNG
   // the same network as SCL:
   #"DI.0.1" := #"DI.a.1";
END_REGION

REGION Network 3
   RUNG wire#powerrail
      Contact( #"DI.a.2" )
      Coil( #"DI.0.2" )
   END_RUNG
   // the same network as SCL:
   #"DI.0.2" := #"DI.a.2";
END_REGION

REGION Network 4
   RUNG wire#powerrail
      Contact( #"DI.a.3" )
      Coil( #"DI.0.3" )
   END_RUNG
   // the same network as SCL:
   #"DI.0.3" := #"DI.a.3";
END_REGION

REGION Network 5
   RUNG wire#powerrail
      Contact( #"DI.a.4" )
      Coil( #"DI.0.4" )
   END_RUNG
   // the same network as SCL:
   #"DI.0.4" := #"DI.a.4";
END_REGION

REGION Network 6
   RUNG wire#powerrail
      Contact( #"DI.a.5" )
      Coil( #"DI.0.5" )
   END_RUNG
   // the same network as SCL:
   #"DI.0.5" := #"DI.a.5";
END_REGION

REGION Network 7
   RUNG wire#powerrail
      Contact( #"DI.a.6" )
      Coil( #"DI.0.6" )
   END_RUNG
   // the same network as SCL:
   #"DI.0.6" := #"DI.a.6";
END_REGION

REGION Network 8
   RUNG wire#powerrail
      Contact( #"DI.a.7" )
      Coil( #"DI.0.7" )
   END_RUNG
   // the same network as SCL:
   #"DI.0.7" := #"DI.a.7";
END_REGION

REGION Network 9
   RUNG wire#powerrail
      I_Contact( #"DI.b.0" )
      Coil( #"DI.1.0" )
   END_RUNG
   // the same network as SCL:
   #"DI.1.0" := NOT #"DI.b.0";
END_REGION

REGION Network 10
   RUNG wire#powerrail
      I_Contact( #"DI.b.1" )
      Coil( #"DI.1.1" )
   END_RUNG
   // the same network as SCL:
   #"DI.1.1" := NOT #"DI.b.1";
END_REGION

REGION Network 11
   RUNG wire#powerrail
      I_Contact( #"DI.b.2" )
      Coil( #"DI.1.2" )
   END_RUNG
   // the same network as SCL:
   #"DI.1.2" := NOT #"DI.b.2";
END_REGION

REGION Network 12
   RUNG wire#powerrail
      I_Contact( #"DI.b.3" )
      Coil( #"DI.1.3" )
   END_RUNG
   // the same network as SCL:
   #"DI.1.3" := NOT #"DI.b.3";
END_REGION

REGION Network 13
   RUNG wire#powerrail
      I_Contact( #"DI.b.4" )
      Coil( #"DI.1.4" )
   END_RUNG
   // the same network as SCL:
   #"DI.1.4" := NOT #"DI.b.4";
END_REGION

REGION Network 14
   RUNG wire#powerrail
      Contact( #"DI.b.5" )
      Coil( #"DI.1.5" )
   END_RUNG
   // the same network as SCL:
   #"DI.1.5" := #"DI.b.5";
END_REGION

REGION Network 15
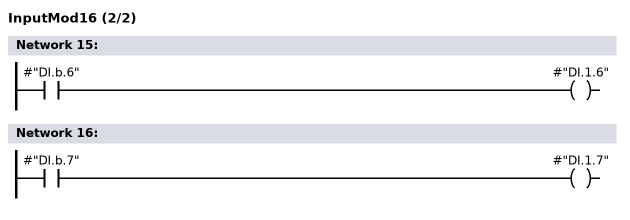
   RUNG wire#powerrail
      Contact( #"DI.b.6" )
      Coil( #"DI.1.6" )
   END_RUNG
   // the same network as SCL:
   #"DI.1.6" := #"DI.b.6";
END_REGION

REGION Network 16
   RUNG wire#powerrail
      Contact( #"DI.b.7" )
      Coil( #"DI.1.7" )
   END_RUNG
   // the same network as SCL:
   #"DI.1.7" := #"DI.b.7";
END_REGION
END_FUNCTION_BLOCK

FUNCTION_BLOCK "OutputMod16"   // FB4, LAD
{ S7_Optimized_Access := 'TRUE' }
VERSION : 0.1
   VAR_INPUT
      "DO.a.0" : Bool;
      "DO.a.1" : Bool;
      "DO.a.2" : Bool;
      "DO.a.3" : Bool;
      "DO.a.4" : Bool;
      "DO.a.5" : Bool;
      "DO.a.6" : Bool;
      "DO.a.7" : Bool;
      "DO.b.0" : Bool;
      "DO.b.1" : Bool;
      "DO.b.2" : Bool;
      "DO.b.3" : Bool;
      "DO.b.4" : Bool;
      "DO.b.5" : Bool;
      "DO.b.6" : Bool;
      "DO.b.7" : Bool;
   END_VAR
   VAR_OUTPUT
      "DO.0.0" : Bool;
      "DO.0.1" : Bool;
      "DO.0.2" : Bool;
      "DO.0.3" : Bool;
      "DO.0.4" : Bool;
      "DO.0.5" : Bool;
      "DO.0.6" : Bool;
      "DO.0.7" : Bool;
      "DO.1.0" : Bool;
      "DO.1.1" : Bool;
      "DO.1.2" : Bool;
      "DO.1.3" : Bool;
      "DO.1.4" : Bool;
      "DO.1.5" : Bool;
      "DO.1.6" : Bool;
      "DO.1.7" : Bool;
   END_VAR
BEGIN

REGION Network 1
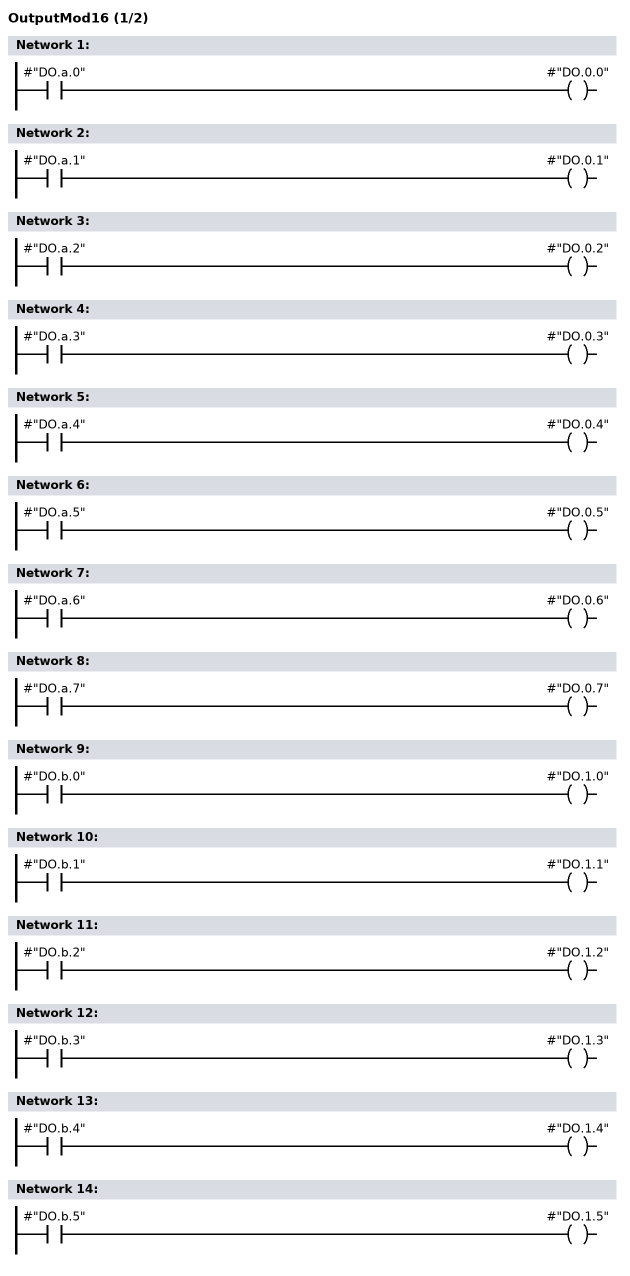
   RUNG wire#powerrail
      Contact( #"DO.a.0" )
      Coil( #"DO.0.0" )
   END_RUNG
   // the same network as SCL:
   #"DO.0.0" := #"DO.a.0";
END_REGION

REGION Network 2
   RUNG wire#powerrail
      Contact( #"DO.a.1" )
      Coil( #"DO.0.1" )
   END_RUNG
   // the same network as SCL:
   #"DO.0.1" := #"DO.a.1";
END_REGION

REGION Network 3
   RUNG wire#powerrail
      Contact( #"DO.a.2" )
      Coil( #"DO.0.2" )
   END_RUNG
   // the same network as SCL:
   #"DO.0.2" := #"DO.a.2";
END_REGION

REGION Network 4
   RUNG wire#powerrail
      Contact( #"DO.a.3" )
      Coil( #"DO.0.3" )
   END_RUNG
   // the same network as SCL:
   #"DO.0.3" := #"DO.a.3";
END_REGION

REGION Network 5
   RUNG wire#powerrail
      Contact( #"DO.a.4" )
      Coil( #"DO.0.4" )
   END_RUNG
   // the same network as SCL:
   #"DO.0.4" := #"DO.a.4";
END_REGION

REGION Network 6
   RUNG wire#powerrail
      Contact( #"DO.a.5" )
      Coil( #"DO.0.5" )
   END_RUNG
   // the same network as SCL:
   #"DO.0.5" := #"DO.a.5";
END_REGION

REGION Network 7
   RUNG wire#powerrail
      Contact( #"DO.a.6" )
      Coil( #"DO.0.6" )
   END_RUNG
   // the same network as SCL:
   #"DO.0.6" := #"DO.a.6";
END_REGION

REGION Network 8
   RUNG wire#powerrail
      Contact( #"DO.a.7" )
      Coil( #"DO.0.7" )
   END_RUNG
   // the same network as SCL:
   #"DO.0.7" := #"DO.a.7";
END_REGION

REGION Network 9
   RUNG wire#powerrail
      Contact( #"DO.b.0" )
      Coil( #"DO.1.0" )
   END_RUNG
   // the same network as SCL:
   #"DO.1.0" := #"DO.b.0";
END_REGION

REGION Network 10
   RUNG wire#powerrail
      Contact( #"DO.b.1" )
      Coil( #"DO.1.1" )
   END_RUNG
   // the same network as SCL:
   #"DO.1.1" := #"DO.b.1";
END_REGION

REGION Network 11
   RUNG wire#powerrail
      Contact( #"DO.b.2" )
      Coil( #"DO.1.2" )
   END_RUNG
   // the same network as SCL:
   #"DO.1.2" := #"DO.b.2";
END_REGION

REGION Network 12
   RUNG wire#powerrail
      Contact( #"DO.b.3" )
      Coil( #"DO.1.3" )
   END_RUNG
   // the same network as SCL:
   #"DO.1.3" := #"DO.b.3";
END_REGION

REGION Network 13
   RUNG wire#powerrail
      Contact( #"DO.b.4" )
      Coil( #"DO.1.4" )
   END_RUNG
   // the same network as SCL:
   #"DO.1.4" := #"DO.b.4";
END_REGION

REGION Network 14
   RUNG wire#powerrail
      Contact( #"DO.b.5" )
      Coil( #"DO.1.5" )
   END_RUNG
   // the same network as SCL:
   #"DO.1.5" := #"DO.b.5";
END_REGION

REGION Network 15
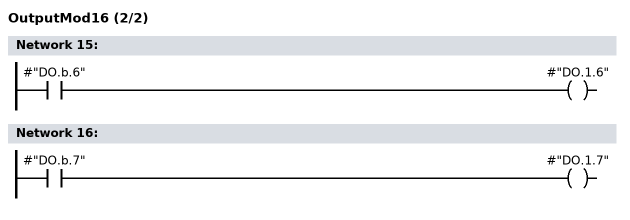
   RUNG wire#powerrail
      Contact( #"DO.b.6" )
      Coil( #"DO.1.6" )
   END_RUNG
   // the same network as SCL:
   #"DO.1.6" := #"DO.b.6";
END_REGION

REGION Network 16
   RUNG wire#powerrail
      Contact( #"DO.b.7" )
      Coil( #"DO.1.7" )
   END_RUNG
   // the same network as SCL:
   #"DO.1.7" := #"DO.b.7";
END_REGION
END_FUNCTION_BLOCK

FUNCTION_BLOCK "NivelTanque"   // FB10, LAD
{ S7_Optimized_Access := 'TRUE' }
VERSION : 0.1
   VAR_INPUT
      EntradaAnalogica : Int;
      Pause : Bool;
      Offset : Real := 500.0;
      Circunferencia : Real := 5.0;
      FirstScan : Bool;
      TempoAtualiza : Time := T#5S;
   END_VAR
   VAR_OUTPUT
      OutKilos : Real;
      OutTon : Real;
   END_VAR
   VAR_IN_OUT
      FatorCorrecao : Real;
   END_VAR
   VAR RETAIN
      OutValor : Real;
      TON_Delay1 : TON_TIME;
      TON_Delay2 : TON_TIME;
      TON_Delay3 : TON_TIME;
      AtualizaLeitura : Bool;
      RaioTanque : Real;
      OutValorCorrigido : Real;
      ValorFisico : Real;
      auxFator : Real;
      CalibraFator : Bool;
      pCalibraFator : Bool;
   END_VAR
   VAR_TEMP
      AUX : Real;
      auxAtualiza : Bool;
   END_VAR
   VAR_TEMP   // added for the SCL form of the ladder/FBD networks
      _w1 : Bool;
   END_VAR
BEGIN

REGION Network 1: Converte o valor da entrada analogica
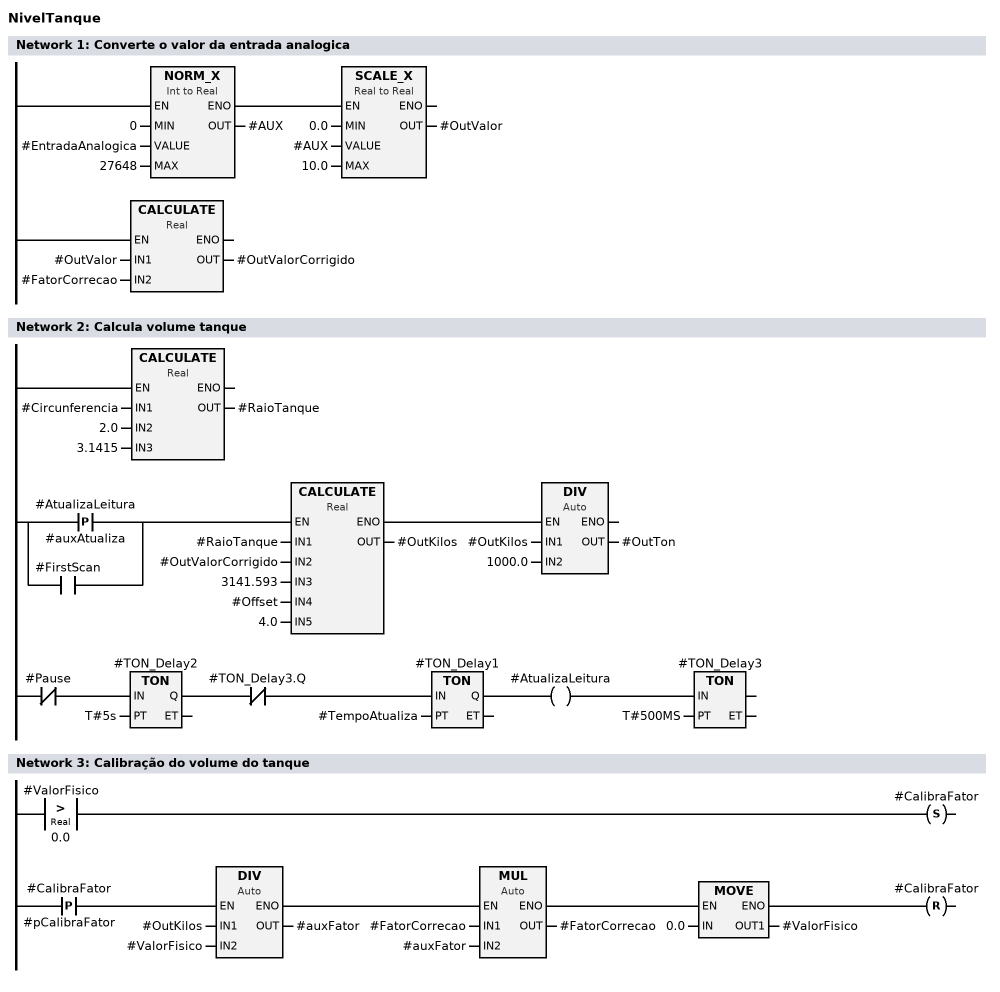
   RUNG wire#powerrail
      { S7_Templates := "[SrcType := Int, DestType := Real]" } Normalize(min := 0, value := #EntradaAnalogica, max := 27648, out => #AUX)
      { S7_Templates := "[SrcType := Real, DestType := Real]" } Scale(min := 0.0, value := #AUX, max := 10.0, out => #OutValor)
   END_RUNG
   RUNG wire#powerrail
      { S7_Templates := "SrcType := Real"; S7_Expression := "(IN1 * IN2)" } Calculate(in1 := #OutValor, in2 := #FatorCorrecao, out => #OutValorCorrigido)
   END_RUNG
   // the same network as SCL:
   #AUX := NORM_X(MIN := 0, VALUE := #EntradaAnalogica, MAX := 27648);
   #OutValor := SCALE_X(MIN := 0.0, VALUE := #AUX, MAX := 10.0);
   #OutValorCorrigido := (#OutValor * #FatorCorrecao);
END_REGION

REGION Network 2: Calcula volume tanque
   #RaioTanque := (#Circunferencia / 2.0 / 3.1415);
   #_w1 := #AtualizaLeitura AND NOT #auxAtualiza;   // rising edge of #AtualizaLeitura
   #auxAtualiza := #AtualizaLeitura;
   IF #_w1 OR #FirstScan THEN
       #OutKilos := (((#RaioTanque * #RaioTanque * #OutValorCorrigido * 3141.593) + #Offset) / 4.0);
       #OutTon := #OutKilos / 1000.0;
   END_IF;
   #TON_Delay2(IN := NOT #Pause, PT := T#5s);   // TON
   #TON_Delay1(IN := #TON_Delay2.Q AND NOT #TON_Delay3.Q, PT := #TempoAtualiza);   // TON
   #AtualizaLeitura := #TON_Delay1.Q;
   #TON_Delay3(IN := #TON_Delay1.Q, PT := T#500MS);   // TON
END_REGION

REGION Network 3: Calibração do volume do tanque
   RUNG wire#powerrail
      { S7_Templates := "SrcType := Real" } GT_Contact(in1 := #ValorFisico, in2 := 0.0)
      S_Coil( #CalibraFator )
   END_RUNG
   RUNG wire#powerrail
      P_Contact(operand := #CalibraFator, bit := #pCalibraFator)
      Div(in1 := #OutKilos, in2 := #ValorFisico, out => #auxFator)
      Mul(in1 := #FatorCorrecao, in2 := #auxFator, out => #FatorCorrecao)
      Move(in := 0.0, out1 => #ValorFisico)
      R_Coil( #CalibraFator )
   END_RUNG
   // the same network as SCL:
   IF #ValorFisico > 0.0 THEN #CalibraFator := TRUE; END_IF;
   #_w1 := #CalibraFator AND NOT #pCalibraFator;   // rising edge of #CalibraFator
   #pCalibraFator := #CalibraFator;
   IF #_w1 THEN
       #auxFator := #OutKilos / #ValorFisico;
       #FatorCorrecao := #FatorCorrecao * #auxFator;
       #ValorFisico := 0.0;
       #CalibraFator := FALSE;
   END_IF;
END_REGION
END_FUNCTION_BLOCK

FUNCTION_BLOCK "SetDbSapi"   // FB15, SCL
{ S7_Optimized_Access := 'TRUE' }
VERSION : 0.1
   VAR_TEMP
      i : Int;
   END_VAR
BEGIN
   FOR #i := 1 TO 200 DO
       "RelatorioSAPI".Hora[#i] := -1;
   END_FOR;

   "RelatorioSAPI".StatusINT := -1;
   "RelatorioSAPI".StatusReal := -1;
END_FUNCTION_BLOCK

FUNCTION_BLOCK "RegistradorMedidor"   // FB99, LAD
{ S7_Optimized_Access := 'TRUE' }
VERSION : 0.1
   VAR_INPUT
      ReadLigado : Bool;
      PulsoMedidor : Bool := false;   // Entrada digital do medidor de pulso
      VolumePulso_ml : Real := 1.0;   // Volume por pulso em mL (ex.: 10.0)
      MedidorEstragado : Bool;
      JanelaTempo_s : Time := T#1MS;   // Janela de cálculo em segundos (ex.: 1.0)
      Filtro : Real := 0.1;   // Filtro exponencial (0.0 a 1.0), ex.: 0.2
      orFlowRate : Real;
   END_VAR
   VAR_OUTPUT
      VolumeAcionamento_L : Real := 0.0;   // Volume total em litros
      DuracaoAcionamento_s : Real;   // Duração do acionamento em segundos
      VazaoFiltrada_Lmin : Real := 0.0;   // Vazão filtrada em litros por minuto
      VazaoFiltrada_Lhora : Real;   // Vazão filtrada em litros por hora
   END_VAR
   VAR_IN_OUT
      VolumeDiario_L : Real;   // Volume dosado no dia em litros
      VolumeTotal_L : LReal;   // Volume totalizar em litros
      DuracaoDiaria_s : Real;   // Tempo ligado no dia em segundos
      DuracaoTotal_s : LReal;   // Tempo ligado no total em segundos
   END_VAR
   VAR RETAIN
      JanelaDone : Bool := false;
      pPulseSignal : Bool;
      TON_TempoJanela : TON_TIME;
      JanelaTempo_ms : DInt;
      Vazao_Lseg : Real;
      temp1 : Real;
      temp2 : Real;
      temp3 : Real;
      Vazao_Lmin : Real := 0.0;   // Vazão instantânea sem filtro
      Vazao_Lhora : Real;   // Vazão instantanea litros
      PulsosJanela : Int;
      VolumePulso_L : Real;
      pClock_10Hz_2 : Bool;
      GravarAcumulado : Bool;
      GravarDiario : Bool;
      GravarTotal : Bool;
      TOF_DelayAcumulado : TOF_TIME;
      TON_DelayZeraAcumulados : TON_TIME;
      TON_DelaySalvaAcumulado : TON_TIME;
      pClock_10Hz_1 : Bool;
      auxFiltro : Real;
      VolumeSeg_L : Real;
      TON_EvitaZerarErrado : TON_TIME;
   END_VAR
   VAR_TEMP   // added for the SCL form of the ladder/FBD networks
      _w1 : Bool;
      _w2 : Bool;
      _w3 : Bool;
      _w4 : Bool;
   END_VAR
BEGIN

REGION Network 1: Contabilização dos pulsos e tempos
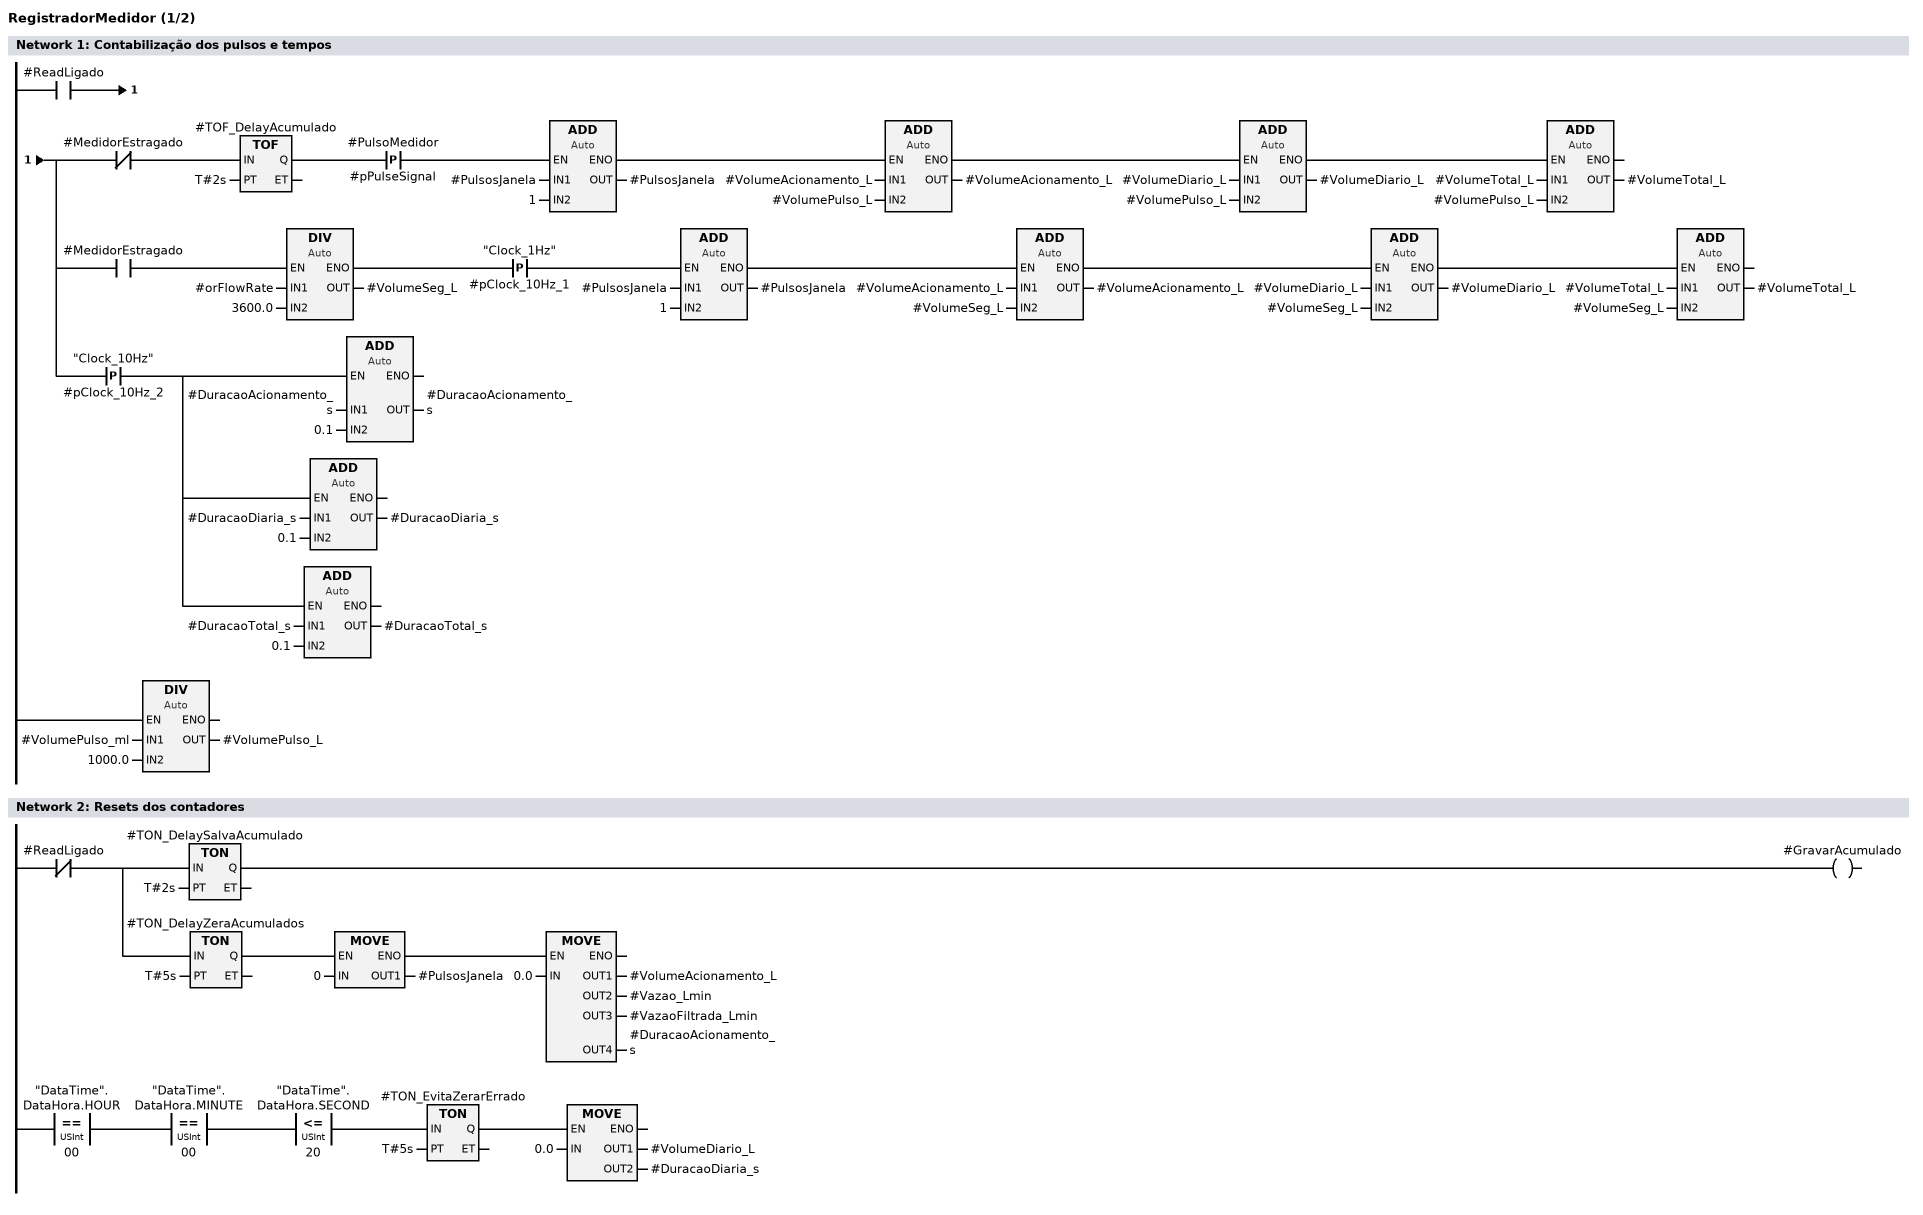
   #TOF_DelayAcumulado(IN := #ReadLigado AND NOT #MedidorEstragado, PT := T#2s);   // TOF
   #_w1 := #TOF_DelayAcumulado.Q AND #PulsoMedidor AND NOT #pPulseSignal;   // rising edge of #PulsoMedidor
   #pPulseSignal := #PulsoMedidor;
   IF #_w1 THEN
       #PulsosJanela := #PulsosJanela + 1;
       #VolumeAcionamento_L := #VolumeAcionamento_L + #VolumePulso_L;
       #VolumeDiario_L := #VolumeDiario_L + #VolumePulso_L;
       #VolumeTotal_L := #VolumeTotal_L + #VolumePulso_L;
   END_IF;
   #_w2 := #ReadLigado AND #MedidorEstragado;
   IF #_w2 THEN #VolumeSeg_L := #orFlowRate / 3600.0; END_IF;
   #_w3 := #_w2 AND "Clock_1Hz" AND NOT #pClock_10Hz_1;   // rising edge of "Clock_1Hz"
   #pClock_10Hz_1 := "Clock_1Hz";
   IF #_w3 THEN
       #PulsosJanela := #PulsosJanela + 1;
       #VolumeAcionamento_L := #VolumeAcionamento_L + #VolumeSeg_L;
       #VolumeDiario_L := #VolumeDiario_L + #VolumeSeg_L;
       #VolumeTotal_L := #VolumeTotal_L + #VolumeSeg_L;
   END_IF;
   #_w4 := #ReadLigado AND "Clock_10Hz" AND NOT #pClock_10Hz_2;   // rising edge of "Clock_10Hz"
   #pClock_10Hz_2 := "Clock_10Hz";
   IF #_w4 THEN
       #DuracaoAcionamento_s := #DuracaoAcionamento_s + 0.1;
       #DuracaoDiaria_s := #DuracaoDiaria_s + 0.1;
       #DuracaoTotal_s := #DuracaoTotal_s + 0.1;
   END_IF;
   #VolumePulso_L := #VolumePulso_ml / 1000.0;
END_REGION

REGION Network 2: Resets dos contadores
   #TON_DelaySalvaAcumulado(IN := NOT #ReadLigado, PT := T#2s);   // TON
   #GravarAcumulado := #TON_DelaySalvaAcumulado.Q;
   #TON_DelayZeraAcumulados(IN := NOT #ReadLigado, PT := T#5s);   // TON
   IF #TON_DelayZeraAcumulados.Q THEN
       #PulsosJanela := 0;
       #VolumeAcionamento_L := 0.0;
       #Vazao_Lmin := 0.0;
       #VazaoFiltrada_Lmin := 0.0;
       #DuracaoAcionamento_s := 0.0;
   END_IF;
   #TON_EvitaZerarErrado(IN := ("DataTime".DataHora.HOUR = 00) AND ("DataTime".DataHora.MINUTE = 00) AND ("DataTime".DataHora.SECOND <= 20),   // TON
                         PT := T#5s);
   IF #TON_EvitaZerarErrado.Q THEN
       #VolumeDiario_L := 0.0;
       #DuracaoDiaria_s := 0.0;
   END_IF;
END_REGION

REGION Network 3: Trigger para os relatorios
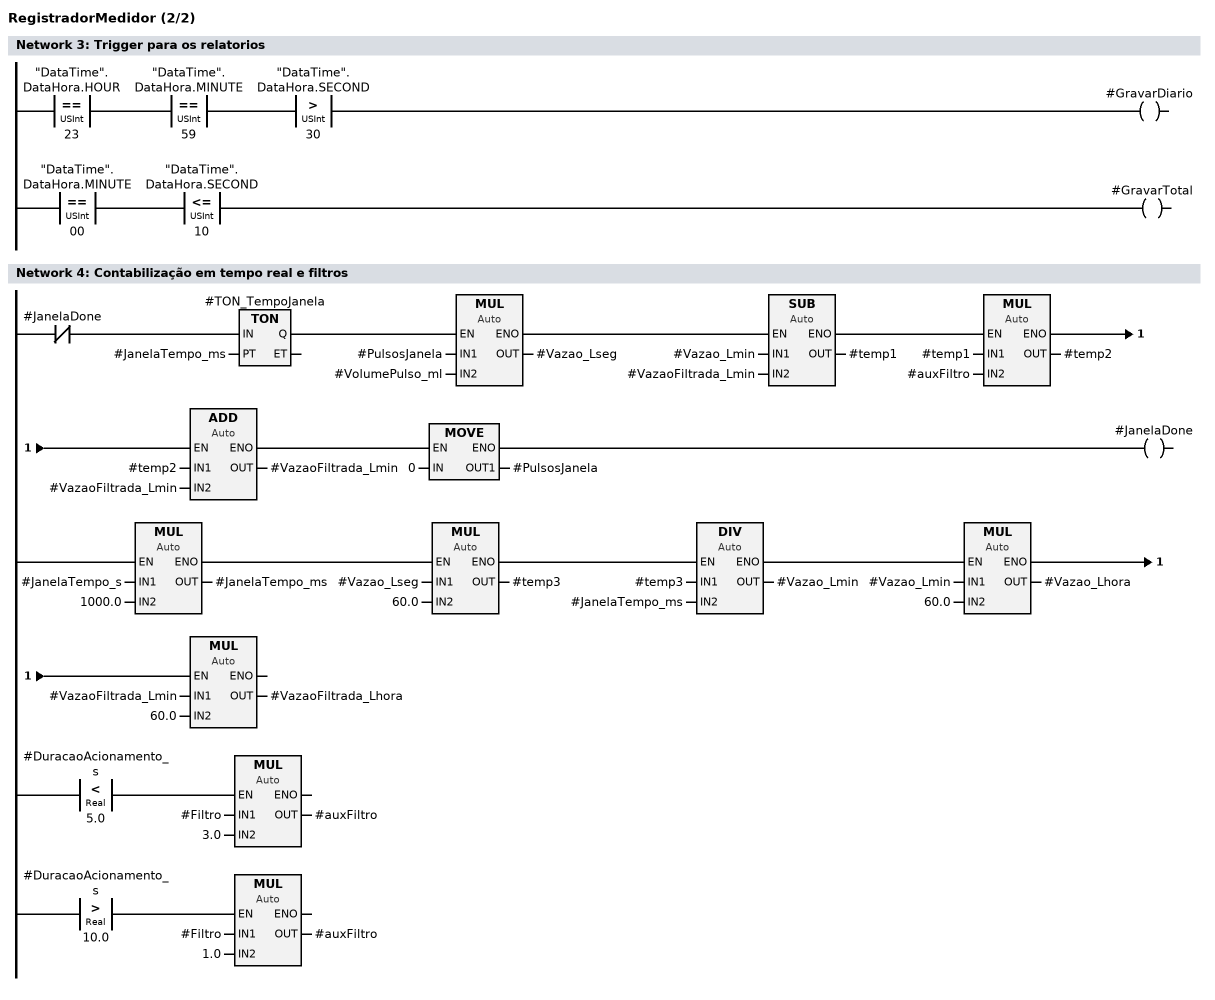
   RUNG wire#powerrail
      { S7_Templates := "SrcType := USInt" } EQ_Contact(in1 := "DataTime".DataHora.HOUR, in2 := 23)
      { S7_Templates := "SrcType := USInt" } EQ_Contact(in1 := "DataTime".DataHora.MINUTE, in2 := 59)
      { S7_Templates := "SrcType := USInt" } GT_Contact(in1 := "DataTime".DataHora.SECOND, in2 := 30)
      Coil( #GravarDiario )
   END_RUNG
   RUNG wire#powerrail
      { S7_Templates := "SrcType := USInt" } EQ_Contact(in1 := "DataTime".DataHora.MINUTE, in2 := 00)
      { S7_Templates := "SrcType := USInt" } LE_Contact(in1 := "DataTime".DataHora.SECOND, in2 := 10)
      Coil( #GravarTotal )
   END_RUNG
   // the same network as SCL:
   #GravarDiario := ("DataTime".DataHora.HOUR = 23) AND ("DataTime".DataHora.MINUTE = 59) AND ("DataTime".DataHora.SECOND > 30);
   #GravarTotal := ("DataTime".DataHora.MINUTE = 00) AND ("DataTime".DataHora.SECOND <= 10);
END_REGION

REGION Network 4: Contabilização em tempo real e filtros
   #TON_TempoJanela(IN := NOT #JanelaDone, PT := #JanelaTempo_ms);   // TON
   IF #TON_TempoJanela.Q THEN
       #Vazao_Lseg := #PulsosJanela * #VolumePulso_ml;
       #temp1 := #Vazao_Lmin - #VazaoFiltrada_Lmin;
       #temp2 := #temp1 * #auxFiltro;
       #VazaoFiltrada_Lmin := #temp2 + #VazaoFiltrada_Lmin;
       #PulsosJanela := 0;
   END_IF;
   #JanelaDone := #TON_TempoJanela.Q;
   #JanelaTempo_ms := #JanelaTempo_s * 1000.0;
   #temp3 := #Vazao_Lseg * 60.0;
   #Vazao_Lmin := #temp3 / #JanelaTempo_ms;
   #Vazao_Lhora := #Vazao_Lmin * 60.0;
   #VazaoFiltrada_Lhora := #VazaoFiltrada_Lmin * 60.0;
   IF #DuracaoAcionamento_s < 5.0 THEN #auxFiltro := #Filtro * 3.0; END_IF;
   IF #DuracaoAcionamento_s > 10.0 THEN #auxFiltro := #Filtro * 1.0; END_IF;
END_REGION
END_FUNCTION_BLOCK

FUNCTION_BLOCK "DosagemCalda2Mist4Inv"   // FB100, LAD
{ S7_Optimized_Access := 'TRUE' }
VERSION : 0.1
   VAR_INPUT
      Clock1Hz : Bool;
      Emergencia : Bool;
      SinalDosagem1 : Bool;
      SinalDosagem2 : Bool;
      RetPesoBalanca1 : Real;
      RetPesoBalanca2 : Real;
      RetValvProd1 : Bool;
      RetValvProd2 : Bool;
      SP_QuantProd1 : Real;
      SP_QuantProd2 : Real;
      SP_QuantAgua1 : Real;
      SP_QuantAgua2 : Real;
      SP_TempoMaxAbastProd1 : Time;
      SP_TempoMaxAbastProd2 : Time;
      SP_TempoMaxAbastAgua1 : Time;
      SP_TempoMaxAbastAgua2 : Time;
      SP_TempoMaxDosagem1 : Time;
      SP_TempoMaxDosagem2 : Time;
      SP_TempMistSeca1 : Time;
      SP_TempMistSeca2 : Time;
      SP_FreqMaxProd1 : Real;
      SP_FreqMaxProd2 : Real;
      SP_FreqMaxAgua1 : Real;
      SP_FreqMaxAgua2 : Real;
      SP_FreqMaxDosagem1 : Real;
      SP_FreqMaxDosagem2 : Real;
      SP_FreqMinProd1 : Real;
      SP_FreqMinProd2 : Real;
      SP_FreqMinAgua1 : Real;
      SP_FreqMinAgua2 : Real;
      SP_FreqMinDosagem1 : Real;
      SP_FreqMinDosagem2 : Real;
      SP_AjusteFinoProd1 : Real;
      SP_AjusteFinoProd2 : Real;
      SP_AjusteFinoAgua1 : Real;
      SP_AjusteFinoAgua2 : Real;
      SP_AjusteFinoDosagem1 : Real;
      SP_AjusteFinoDosagem2 : Real;
      SP_CorteProd1 : Real;
      SP_CorteProd2 : Real;
      SP_CorteAgua1 : Real;
      SP_CorteAgua2 : Real;
      SP_CorteDosagem1 : Real;
      SP_CorteDosagem2 : Real;
      SP_Transbordo1 : Real;
      SP_Transbordo2 : Real;
      ReadLigadoProd : Bool;
      ReadLigadoAgua : Bool;
      ReadLigadoDosagem1 : Bool;
      ReadLigadoDosagem2 : Bool;
      IN_FalhaBomba1 : Bool;
      IN_FalhaBomba2 : Bool;
      IN_FalhaBomba3 : Bool;
      IN_FalhaBomba4 : Bool;
      ProdFim1 : Bool;
      ProdFim2 : Bool;
      AguaFim1 : Bool;
      AguaFim2 : Bool;
      IniciaAbast1 : Bool;
      IniciaAbast2 : Bool;
   END_VAR
   VAR_OUTPUT
      LigarBomba1 : Bool;
      LigarBomba2 : Bool;
      LigarBomba3 : Bool;
      LigarBomba4 : Bool;
      AcionaValvProd1 : Bool;
      AcionaValvProd2 : Bool;
      AcionaValvAgua1 : Bool;
      AcionaValvAgua2 : Bool;
      AcionaValvDos1 : Bool;
      AcionaValvDos2 : Bool;
      FreqAtual1 : Real;
      FreqAtual2 : Real;
      FreqAtual3 : Real;
      FreqAtual4 : Real;
      FalhaBomba1 : Bool;
      FalhaBomba2 : Bool;
      FalhaBomba3 : Bool;
      FalhaBomba4 : Bool;
   END_VAR
   VAR_IN_OUT
      DosadoDiarioProduto1 : Real;
      DosadoDiarioProduto2 : Real;
      DosadoDiarioAgua1 : Real;
      DosadoDiarioAgua2 : Real;
      DosadoDiarioCalda1 : Real;
      DosadoDiarioCalda2 : Real;
      DosadoTotalProduto1 : Real;
      DosadoTotalProduto2 : Real;
      DosadoTotalAgua1 : Real;
      DosadoTotalAgua2 : Real;
      DosadoTotalCalda1 : Real;
      DosadoTotalCalda2 : Real;
      DuracaoDiariaProduto1 : DInt;
      DuracaoDiariaProduto2 : DInt;
      DuracaoDiariaAgua1 : DInt;
      DuracaoDiariaAgua2 : DInt;
      DuracaoDiariaCalda1 : DInt;
      DuracaoDiariaCalda2 : DInt;
      DuracaoTotalProduto1 : DInt;
      DuracaoTotalProduto2 : DInt;
      DuracaoTotalAgua1 : DInt;
      DuracaoTotalAgua2 : DInt;
      DuracaoTotalCalda1 : DInt;
      DuracaoTotalCalda2 : DInt;
   END_VAR
   VAR RETAIN
      TON_EstabilizaBalancaProduto1 : TON_TIME;
      TON_EstabilizaBalancaProduto2 : TON_TIME;
      TON_EstabilizaBalancaAgua1 : TON_TIME;
      TON_EstabilizaBalancaAgua2 : TON_TIME;
      AcionaFreqMinProd1 : Bool;
      AcionaFreqMinProd2 : Bool;
      AcionaFreqMinAgua1 : Bool;
      AcionaFreqMinAgua2 : Bool;
      AcionaFreqMinDosagem1 : Bool;
      AcionaFreqMinDosagem2 : Bool;
      ProdutoFinalizado1 : Bool;
      ProdutoFinalizado2 : Bool;
      auxPesoBal1 : Real;
      auxPesoBal2 : Real;
      QuantAlvoProd1 : Real;
      QuantAlvoProd2 : Real;
      BalancaVazia1 : Bool;
      BalancaVazia2 : Bool;
      AguaFinalizada1 : Bool;
      AguaFinalizada2 : Bool;
      QuantAlvoAgua1 : Real;
      QuantAlvoAgua2 : Real;
      auxPulsoSinalDosagem1 : Bool;
      auxPulsoSinalDosagem2 : Bool;
      TON_MisturaSeca1 : TON_TIME;
      TON_MisturaSeca2 : TON_TIME;
      auxSetSinalDosagem1 : Bool;
      auxSetSinalDosagem2 : Bool;
      HabilitadoDosagem1 : Bool;
      HabilitadoDosagem2 : Bool;
      QuantAjusteProd1 : Real;
      QuantAjusteProd2 : Real;
      QuantAjusteAgua1 : Real;
      QuantAjusteAgua2 : Real;
      auxPulsoBatidaFinalizada1 : Bool;
      auxPulsoBatidaFinalizada2 : Bool;
      auxPulsoLigarBombaProd1 : Bool;
      auxPulsoLigarBombaProd2 : Bool;
      auxPulsoLigarBombaAgua1 : Bool;
      auxPulsoLigarBombaAgua2 : Bool;
      auxPulsoLigarBombaDosagem1 : Bool;
      auxPulsoLigarBombaDosagem2 : Bool;
      TON_TempoMaxDos1 : TON_TIME;
      TON_TempoMaxDos2 : TON_TIME;
      TON_TempoMaxAbastProd1 : TON_TIME;
      TON_TempoMaxAbastProd2 : TON_TIME;
      TON_TempoMaxAbastAgua1 : TON_TIME;
      TON_TempoMaxAbastAgua2 : TON_TIME;
      auxTempoMisturaSeca1 : Time;
      auxTempoMisturaSeca2 : Time;
      auxTempoMaxAbastProd1 : DInt;
      auxTempoMaxAbastProd2 : DInt;
      auxTempoMaxAbastAgua1 : DInt;
      auxTempoMaxAbastAgua2 : DInt;
      auxTempoMaxDosagem1 : DInt;
      auxTempoMaxDosagem2 : DInt;
      auxTempoMax1 : DInt;
      auxTempoMax2 : DInt;
      TON_ResetSinalFabrica1 : TON_TIME;
      TON_ResetSinalFabrica2 : TON_TIME;
      TOF_RegistraPesoCalda1 : TOF_TIME;
      TOF_RegistraPesoCalda2 : TOF_TIME;
      TOF_RegistraPesoProd1 : TOF_TIME;
      TOF_RegistraPesoProd2 : TOF_TIME;
      TOF_RegistraPesoAgua1 : TOF_TIME;
      TOF_RegistraPesoAgua2 : TOF_TIME;
      TON_FalhaRetornoBomba1 : TON_TIME;
      TON_FalhaRetornoBomba2 : TON_TIME;
      TON_FalhaRetornoBomba3 : TON_TIME;
      TON_FalhaRetornoBomba4 : TON_TIME;
      auxTempoMisturaSecaDecorrido1 : DInt;
      auxTempoMisturaSecaDecorrido2 : DInt;
      auxPulsoClock1HZ : Array[0..10] of Bool;
      auxTempoTotal1 : DInt;
      auxTempoTotal2 : DInt;
      TOF_BatidaFinalizada1 : TOF_TIME;
      TOF_BatidaFinalizada2 : TOF_TIME;
      SistemaHabilitado1 : Bool;
      SistemaHabilitado2 : Bool;
      Manual1 : Bool;
      Manual2 : Bool;
      Manual3 : Bool;
      Manual4 : Bool;
      LigaManualProd1 : Bool;
      LigaManualProd2 : Bool;
      LigaManualAgua1 : Bool;
      LigaManualAgua2 : Bool;
      LigaManualDos1 : Bool;
      LigaManualDos2 : Bool;
      Manutencao1 : Bool;
      Manutencao2 : Bool;
      Manutencao3 : Bool;
      Manutencao4 : Bool;
      GravarDiario : Bool;
      GravarTotalizador : Bool;
      DuracaoBatProduto1 : DInt;
      DuracaoBatProduto2 : DInt;
      DuracaoBatAgua1 : DInt;
      DuracaoBatAgua2 : DInt;
      DuracaoBatCalda1 : DInt;
      DuracaoBatCalda2 : DInt;
      DosadoBatProduto1 : Real;
      DosadoBatProduto2 : Real;
      DosadoBatAgua1 : Real;
      DosadoBatAgua2 : Real;
      DosadoBatCalda1 : Real;
      DosadoBatCalda2 : Real;
      TempoMaxDosRestanteMS1 : DInt;
      TempoMaxDosRestanteMS2 : DInt;
      TempoMaxDosRestanteSeg1 : DInt;
      TempoMaxDosRestanteSeg2 : DInt;
      FalhaTempoMaxAbastProd1 : Bool;
      FalhaTempoMaxAbastProd2 : Bool;
      FalhaTempoMaxAbastAgua1 : Bool;
      FalhaTempoMaxAbastAgua2 : Bool;
      FalhaTempoMax1 : Bool;
      FalhaTempoMax2 : Bool;
      FalhaTransbordo1 : Bool;
      FalhaTransbordo2 : Bool;
      BatidaFinalizada1 : Bool;
      BatidaFinalizada2 : Bool;
      CaldaFinalizada1 : Bool;
      CaldaFinalizada2 : Bool;
      StatusBomba1 : Int;
      StatusBomba2 : Int;
      StatusBomba3 : Int;
      StatusBomba4 : Int;
      StatusIcone1 : Int;
      StatusIcone2 : Int;
      StatusIcone3 : Int;
      StatusIcone4 : Int;
      AbastecendoProd1 : Bool;
      AbastecendoProd2 : Bool;
      AbastecendoAgua1 : Bool;
      AbastecendoAgua2 : Bool;
      DosadoProdIHM : Real;
      DosadoAguaIHM : Real;
      DuracaoProdIHM : DInt;
      DuracaoAguaIHM : DInt;
      auxLigaBomba3 : Bool;
      auxLigaBomba4 : Bool;
      FalhaRetornoBomba1 : Bool;
      FalhaRetornoBomba2 : Bool;
      FalhaRetornoBomba3 : Bool;
      FalhaRetornoBomba4 : Bool;
      GravarBatelada1 : Bool;
      TON_DelayGravaBatelada2 : TON_TIME;
      TON_DelayGravaBatelada1 : TON_TIME;
      GravarBatelada2 : Bool;
      TON_FalhaRetornoValvProd1 : TON_TIME;
      FalhaValvProd1 : Bool;
      TON_FalhaRetornoValvProd2 : TON_TIME;
      FalhaValvProd2 : Bool;
   END_VAR
   VAR_TEMP   // added for the SCL form of the ladder/FBD networks
      _w1 : Bool;
      _w2 : Bool;
      _w3 : Bool;
      _w4 : Bool;
      _w5 : Bool;
      _w6 : Bool;
   END_VAR
BEGIN

REGION Network 1: Prepara calda (Produto 1)
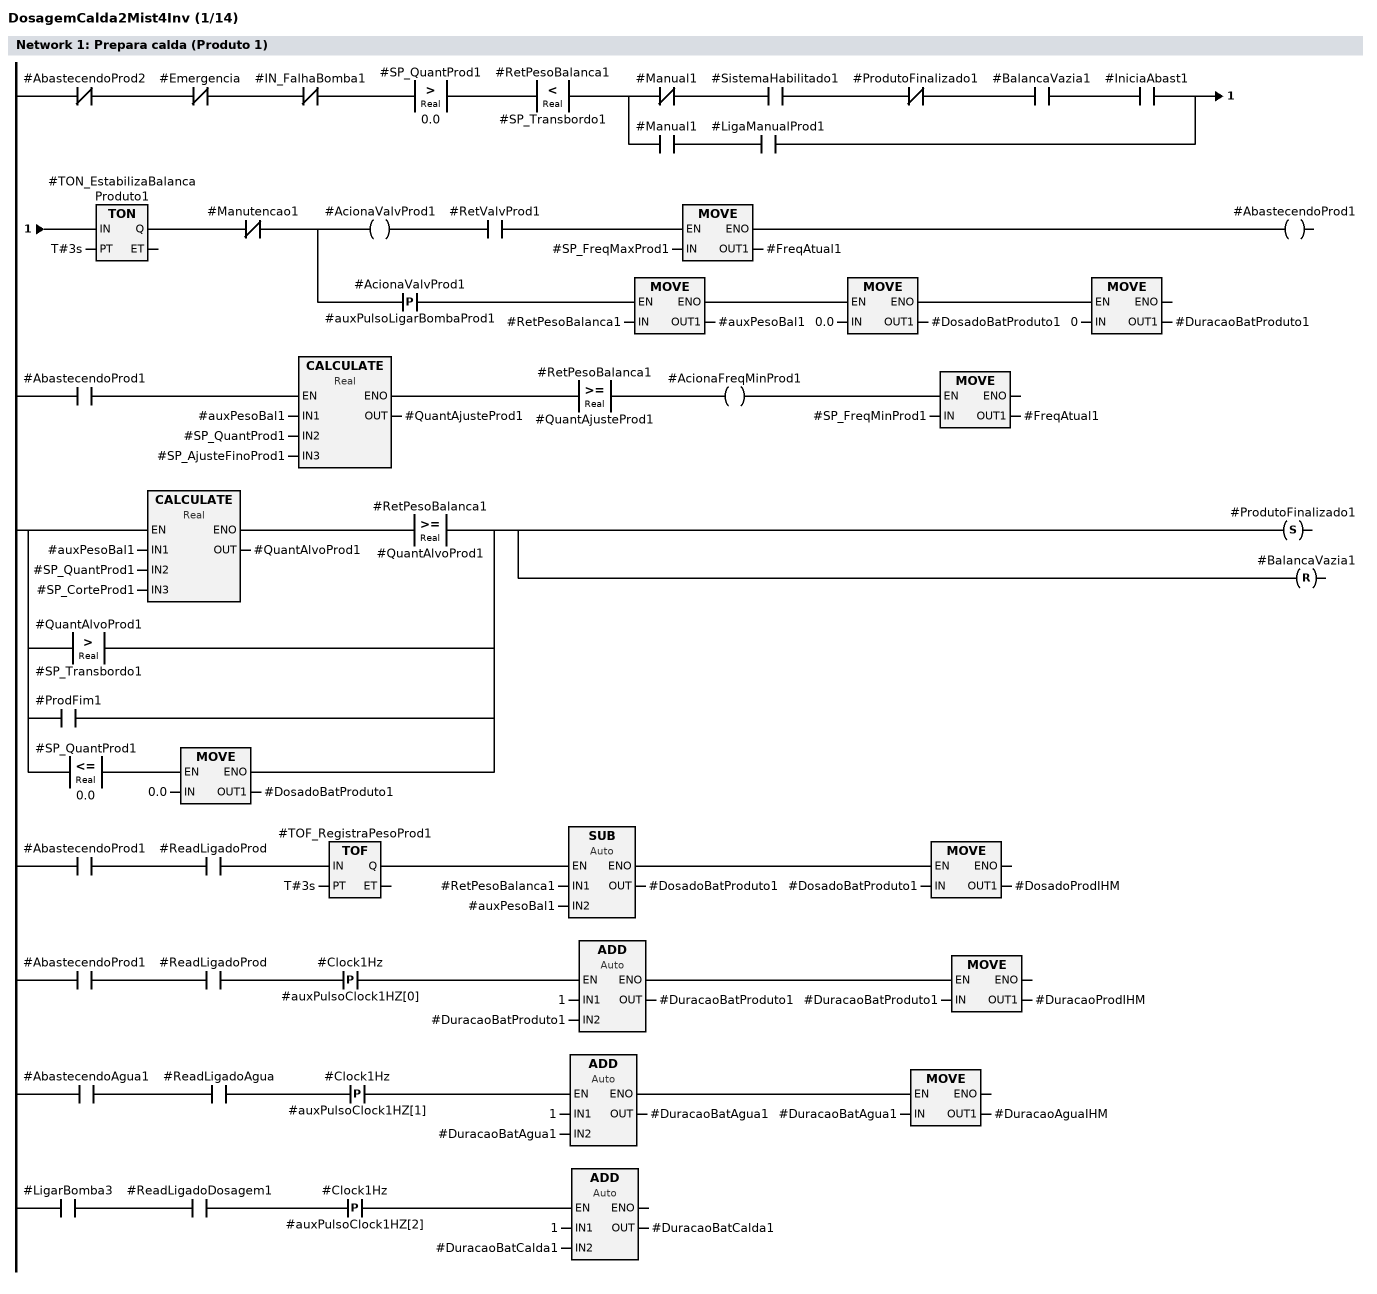
   #TON_EstabilizaBalancaProduto1(IN := NOT #AbastecendoProd2 AND NOT #Emergencia AND NOT #IN_FalhaBomba1 AND (#SP_QuantProd1 > 0.0) AND (#RetPesoBalanca1 < #SP_Transbordo1) AND ((NOT #Manual1 AND #SistemaHabilitado1 AND NOT #ProdutoFinalizado1 AND #BalancaVazia1 AND #IniciaAbast1) OR (#Manual1 AND #LigaManualProd1)),   // TON
                           PT := T#3s);
   #AcionaValvProd1 := #TON_EstabilizaBalancaProduto1.Q AND NOT #Manutencao1;
   #_w1 := #AcionaValvProd1 AND #RetValvProd1;
   IF #_w1 THEN #FreqAtual1 := #SP_FreqMaxProd1; END_IF;
   #AbastecendoProd1 := #_w1;
   #_w2 := #AcionaValvProd1 AND #AcionaValvProd1 AND NOT #auxPulsoLigarBombaProd1;   // rising edge of #AcionaValvProd1
   #auxPulsoLigarBombaProd1 := #AcionaValvProd1;
   IF #_w2 THEN
       #auxPesoBal1 := #RetPesoBalanca1;
       #DosadoBatProduto1 := 0.0;
       #DuracaoBatProduto1 := 0;
   END_IF;
   IF #AbastecendoProd1 THEN
       #QuantAjusteProd1 := (#auxPesoBal1 + #SP_QuantProd1 - #SP_AjusteFinoProd1);
   END_IF;
   #AcionaFreqMinProd1 := #AbastecendoProd1 AND (#RetPesoBalanca1 >= #QuantAjusteProd1);
   IF #AcionaFreqMinProd1 THEN #FreqAtual1 := #SP_FreqMinProd1; END_IF;
   #QuantAlvoProd1 := (#auxPesoBal1 + #SP_QuantProd1 - #SP_CorteProd1);
   #_w3 := #SP_QuantProd1 <= 0.0;
   IF #_w3 THEN #DosadoBatProduto1 := 0.0; END_IF;
   IF (#RetPesoBalanca1 >= #QuantAlvoProd1) OR (#QuantAlvoProd1 > #SP_Transbordo1) OR #ProdFim1 OR #_w3 THEN
       #ProdutoFinalizado1 := TRUE;
       #BalancaVazia1 := FALSE;
   END_IF;
   #TOF_RegistraPesoProd1(IN := #AbastecendoProd1 AND #ReadLigadoProd, PT := T#3s);   // TOF
   IF #TOF_RegistraPesoProd1.Q THEN
       #DosadoBatProduto1 := #RetPesoBalanca1 - #auxPesoBal1;
       #DosadoProdIHM := #DosadoBatProduto1;
   END_IF;
   #_w4 := #AbastecendoProd1 AND #ReadLigadoProd AND #Clock1Hz AND NOT #auxPulsoClock1HZ[0];   // rising edge of #Clock1Hz
   #auxPulsoClock1HZ[0] := #Clock1Hz;
   IF #_w4 THEN
       #DuracaoBatProduto1 := 1 + #DuracaoBatProduto1;
       #DuracaoProdIHM := #DuracaoBatProduto1;
   END_IF;
   #_w5 := #AbastecendoAgua1 AND #ReadLigadoAgua AND #Clock1Hz AND NOT #auxPulsoClock1HZ[1];   // rising edge of #Clock1Hz
   #auxPulsoClock1HZ[1] := #Clock1Hz;
   IF #_w5 THEN
       #DuracaoBatAgua1 := 1 + #DuracaoBatAgua1;
       #DuracaoAguaIHM := #DuracaoBatAgua1;
   END_IF;
   #_w6 := #LigarBomba3 AND #ReadLigadoDosagem1 AND #Clock1Hz AND NOT #auxPulsoClock1HZ[2];   // rising edge of #Clock1Hz
   #auxPulsoClock1HZ[2] := #Clock1Hz;
   IF #_w6 THEN #DuracaoBatCalda1 := 1 + #DuracaoBatCalda1; END_IF;
END_REGION

REGION Network 2: Prepara calda (Produto 2)
